// TIA Portal V20 program export: 0 tag tables, 0 data types, 6 data blocks, 13 code blocks (in call order from the OBs), 34 instance data blocks

DATA_BLOCK "DB_Bad_Konfig"   // DB8
{ S7_Optimized_Access := 'TRUE' }
VERSION : 0.5
// stored: AutoNumber true, DBAccessibleFromOPCUA true, DBAccessibleFromWebserver true, IsOnlyStoredInLoadMemory false, IsRetainMemResEnabled false, IsWriteProtectedInAS false, MemoryReserve 100
   VAR
      Bad_Konfig : Array[1.."c_Anzahl_Bad"] of "UDT_Bad_Konfig";
   END_VAR
BEGIN
   Bad_Konfig[7..8].Ausstattung.HatHeizung_1 := TRUE;
   Bad_Konfig[12].Ausstattung.HatHeizung_1 := TRUE;
   Bad_Konfig[25].Ausstattung.HatHeizung_1 := TRUE;
   Bad_Konfig[36].Ausstattung.HatHeizung_1 := TRUE;
   Bad_Konfig[40].Ausstattung.HatHeizung_1 := TRUE;
   Bad_Konfig[46].Ausstattung.HatHeizung_1 := TRUE;
   Bad_Konfig[25].Ausstattung.HatHeizung_2 := TRUE;
   Bad_Konfig[8].Ausstattung.HatPumpe := TRUE;
   Bad_Konfig[12].Ausstattung.HatPumpe := TRUE;
   Bad_Konfig[14].Ausstattung.HatPumpe := TRUE;
   Bad_Konfig[18..19].Ausstattung.HatPumpe := TRUE;
   Bad_Konfig[21].Ausstattung.HatPumpe := TRUE;
   Bad_Konfig[25..26].Ausstattung.HatPumpe := TRUE;
   Bad_Konfig[31].Ausstattung.HatPumpe := TRUE;
   Bad_Konfig[41].Ausstattung.HatPumpe := TRUE;
   Bad_Konfig[45].Ausstattung.HatPumpe := TRUE;
   Bad_Konfig[25].Ausstattung.HatPumpe_FU := TRUE;
   Bad_Konfig[25].Ausstattung.HatWarenbewegung_X := TRUE;
   Bad_Konfig[25].Ausstattung.HatWarenbewegung_Y := TRUE;
   Bad_Konfig[8].Ausstattung.HatUltraschall := TRUE;
   Bad_Konfig[12].Ausstattung.HatUltraschall := TRUE;
   Bad_Konfig[31].Ausstattung.HatGleichrichter := TRUE;
   Bad_Konfig[36].Ausstattung.HatGleichrichter := TRUE;
   Bad_Konfig[40].Ausstattung.HatGleichrichter := TRUE;
   Bad_Konfig[7..8].Ausstattung.HatNiveau := TRUE;
   Bad_Konfig[12].Ausstattung.HatNiveau := TRUE;
   Bad_Konfig[25].Ausstattung.HatNiveau := TRUE;
   Bad_Konfig[36].Ausstattung.HatNiveau := TRUE;
   Bad_Konfig[40].Ausstattung.HatNiveau := TRUE;
   Bad_Konfig[46].Ausstattung.HatNiveau := TRUE;
   Bad_Konfig[1].WT[1..3].Auftragsindex := -1;
   Bad_Konfig[2].WT[1..3].Auftragsindex := -1;
   Bad_Konfig[3].WT[1..3].Auftragsindex := -1;
   Bad_Konfig[4].WT[1..3].Auftragsindex := -1;
   Bad_Konfig[5].WT[1..3].Auftragsindex := -1;
   Bad_Konfig[6].WT[1..3].Auftragsindex := -1;
   Bad_Konfig[7].WT[1..3].Auftragsindex := -1;
   Bad_Konfig[8].WT[1..3].Auftragsindex := -1;
   Bad_Konfig[9].WT[1..3].Auftragsindex := -1;
   Bad_Konfig[10].WT[1..3].Auftragsindex := -1;
   Bad_Konfig[11].WT[1..3].Auftragsindex := -1;
   Bad_Konfig[12].WT[1..3].Auftragsindex := -1;
   Bad_Konfig[13].WT[1..3].Auftragsindex := -1;
   Bad_Konfig[14].WT[1..3].Auftragsindex := -1;
   Bad_Konfig[15].WT[1..3].Auftragsindex := -1;
   Bad_Konfig[16].WT[1..3].Auftragsindex := -1;
   Bad_Konfig[17].WT[1..3].Auftragsindex := -1;
   Bad_Konfig[18].WT[1..3].Auftragsindex := -1;
   Bad_Konfig[19].WT[1..3].Auftragsindex := -1;
   Bad_Konfig[20].WT[1..3].Auftragsindex := -1;
   Bad_Konfig[21].WT[1..3].Auftragsindex := -1;
   Bad_Konfig[22].WT[1..3].Auftragsindex := -1;
   Bad_Konfig[23].WT[1..3].Auftragsindex := -1;
   Bad_Konfig[24].WT[1..3].Auftragsindex := -1;
   Bad_Konfig[25].WT[1..3].Auftragsindex := -1;
   Bad_Konfig[26].WT[1..3].Auftragsindex := -1;
   Bad_Konfig[27].WT[1..3].Auftragsindex := -1;
   Bad_Konfig[28].WT[1..3].Auftragsindex := -1;
   Bad_Konfig[29].WT[1..3].Auftragsindex := -1;
   Bad_Konfig[30].WT[1..3].Auftragsindex := -1;
   Bad_Konfig[31].WT[1..3].Auftragsindex := -1;
   Bad_Konfig[32].WT[1..3].Auftragsindex := -1;
   Bad_Konfig[33].WT[1..3].Auftragsindex := -1;
   Bad_Konfig[34].WT[1..3].Auftragsindex := -1;
   Bad_Konfig[35].WT[1..3].Auftragsindex := -1;
   Bad_Konfig[36].WT[1..3].Auftragsindex := -1;
   Bad_Konfig[37].WT[1..3].Auftragsindex := -1;
   Bad_Konfig[38].WT[1..3].Auftragsindex := -1;
   Bad_Konfig[39].WT[1..3].Auftragsindex := -1;
   Bad_Konfig[40].WT[1..3].Auftragsindex := -1;
   Bad_Konfig[41].WT[1..3].Auftragsindex := -1;
   Bad_Konfig[42].WT[1..3].Auftragsindex := -1;
   Bad_Konfig[43].WT[1..3].Auftragsindex := -1;
   Bad_Konfig[44].WT[1..3].Auftragsindex := -1;
   Bad_Konfig[45].WT[1..3].Auftragsindex := -1;
   Bad_Konfig[46].WT[1..3].Auftragsindex := -1;
   Bad_Konfig[47].WT[1..3].Auftragsindex := -1;
   Bad_Konfig[1].WT[1..3].SchrittIndex := -1;
   Bad_Konfig[2].WT[1..3].SchrittIndex := -1;
   Bad_Konfig[3].WT[1..3].SchrittIndex := -1;
   Bad_Konfig[4].WT[1..3].SchrittIndex := -1;
   Bad_Konfig[5].WT[1..3].SchrittIndex := -1;
   Bad_Konfig[6].WT[1..3].SchrittIndex := -1;
   Bad_Konfig[7].WT[1..3].SchrittIndex := -1;
   Bad_Konfig[8].WT[1..3].SchrittIndex := -1;
   Bad_Konfig[9].WT[1..3].SchrittIndex := -1;
   Bad_Konfig[10].WT[1..3].SchrittIndex := -1;
   Bad_Konfig[11].WT[1..3].SchrittIndex := -1;
   Bad_Konfig[12].WT[1..3].SchrittIndex := -1;
   Bad_Konfig[13].WT[1..3].SchrittIndex := -1;
   Bad_Konfig[14].WT[1..3].SchrittIndex := -1;
   Bad_Konfig[15].WT[1..3].SchrittIndex := -1;
   Bad_Konfig[16].WT[1..3].SchrittIndex := -1;
   Bad_Konfig[17].WT[1..3].SchrittIndex := -1;
   Bad_Konfig[18].WT[1..3].SchrittIndex := -1;
   Bad_Konfig[19].WT[1..3].SchrittIndex := -1;
   Bad_Konfig[20].WT[1..3].SchrittIndex := -1;
   Bad_Konfig[21].WT[1..3].SchrittIndex := -1;
   Bad_Konfig[22].WT[1..3].SchrittIndex := -1;
   Bad_Konfig[23].WT[1..3].SchrittIndex := -1;
   Bad_Konfig[24].WT[1..3].SchrittIndex := -1;
   Bad_Konfig[25].WT[1..3].SchrittIndex := -1;
   Bad_Konfig[26].WT[1..3].SchrittIndex := -1;
   Bad_Konfig[27].WT[1..3].SchrittIndex := -1;
   Bad_Konfig[28].WT[1..3].SchrittIndex := -1;
   Bad_Konfig[29].WT[1..3].SchrittIndex := -1;
   Bad_Konfig[30].WT[1..3].SchrittIndex := -1;
   Bad_Konfig[31].WT[1..3].SchrittIndex := -1;
   Bad_Konfig[32].WT[1..3].SchrittIndex := -1;
   Bad_Konfig[33].WT[1..3].SchrittIndex := -1;
   Bad_Konfig[34].WT[1..3].SchrittIndex := -1;
   Bad_Konfig[35].WT[1..3].SchrittIndex := -1;
   Bad_Konfig[36].WT[1..3].SchrittIndex := -1;
   Bad_Konfig[37].WT[1..3].SchrittIndex := -1;
   Bad_Konfig[38].WT[1..3].SchrittIndex := -1;
   Bad_Konfig[39].WT[1..3].SchrittIndex := -1;
   Bad_Konfig[40].WT[1..3].SchrittIndex := -1;
   Bad_Konfig[41].WT[1..3].SchrittIndex := -1;
   Bad_Konfig[42].WT[1..3].SchrittIndex := -1;
   Bad_Konfig[43].WT[1..3].SchrittIndex := -1;
   Bad_Konfig[44].WT[1..3].SchrittIndex := -1;
   Bad_Konfig[45].WT[1..3].SchrittIndex := -1;
   Bad_Konfig[46].WT[1..3].SchrittIndex := -1;
   Bad_Konfig[47].WT[1..3].SchrittIndex := -1;
END_DATA_BLOCK

DATA_BLOCK "DB_HMI"   // DB4
{ S7_Optimized_Access := 'TRUE' }
VERSION : 0.1
// stored: AutoNumber true, DBAccessibleFromOPCUA true, DBAccessibleFromWebserver true, IsOnlyStoredInLoadMemory false, IsRetainMemResEnabled false, IsWriteProtectedInAS false, MemoryReserve 100
   VAR
      Benutzerverwaltung_User_Daten { S7_SetPoint := 'True'} : "UDT_Benutzer";
      Benutzerverwaltung_User_create { S7_SetPoint := 'True'} : Bool;
      Benutzerverwaltung_User_update : Bool;
      Benutzerverwaltung_User_delete : Bool;
      Benutzerverwaltung_Freigaben_Prozessgruppen_User_change : Bool;
      Benutzerverwaltung_Status : Int;
      Benutzerverwaltung_Freigabe_Prozessgruppen_User_ID_ausgewählt : Int;
      Benutzerverwaltung_Freigabe_Prozessgruppen_Prozessgruppen : Array[1.."c_Prozessgruppen"] of Bool;
      Benutzerverwaltung_Login_Name : String;
      Benutzerverwaltung_Login_Passwort : String;
      Benutzerverwaltung_Login_Loginbutton : Bool;
      Benutzerverwaltung_Login_Logoutbutton : Bool;
      Benutzerverwaltung_Login_Login_Ok : Bool;
      Prozessparameter_Status : Int;
      Prozessparameter_Prozessgruppen_save : Bool;
      Prozessparameter_Prozessgruppen_Prozessgruppe : "UDT_Prozessgruppen";
      Prozessparameter_Artikel_add { S7_SetPoint := 'True'} : "UDT_Artikel";
      Prozessparameter_Artikel_save { S7_SetPoint := 'True'} : Bool;
      Prozessparameter_Artikel_delete : Bool;
      Prozessparameter_Artikel_assign : Bool;
      Prozessparameter_Artikel_remove : Bool;
      "Prozessparameter_Prozessgruppe_ID_assign/remove" : Int;
      "Prozessparameter_Artikel_ID_assign/remove" : Int;
      Angewähltes_Bad : USInt;
      Handbetrieb { S7_SetPoint := 'True'} : "UDT_Handbetrieb";
   END_VAR
BEGIN
END_DATA_BLOCK

DATA_BLOCK "DB_CPU_to_IPC"   // DB3
{ S7_Optimized_Access := 'TRUE' }
VERSION : 0.2
// stored: AutoNumber true, DBAccessibleFromOPCUA true, DBAccessibleFromWebserver true, IsOnlyStoredInLoadMemory false, IsRetainMemResEnabled false, IsWriteProtectedInAS false, MemoryReserve 100
   VAR
      Bad : Array[1.."c_Anzahl_Bad"] of "UDT_Bad_Rueckmeldung";
      Not_Halt_Aktiv : Bool;
      Not_Aus_OK : Bool;
      Auftrag_Abgeschlossen : Array[0..9] of Bool;
   END_VAR
BEGIN
END_DATA_BLOCK

DATA_BLOCK "DB_Fehlermeldungen"   // DB39
{ S7_Optimized_Access := 'TRUE' }
VERSION : 0.2
// FI-Schutz ausgeloest (Heizungen)
// stored: AutoNumber true, DBAccessibleFromOPCUA true, DBAccessibleFromWebserver true, IsOnlyStoredInLoadMemory false, IsRetainMemResEnabled false, IsWriteProtectedInAS false, MemoryReserve 100
   VAR
      FI_Heizung_Bad_7 : Bool;   // 1 - FI-Schutz 200F1 Heizung Bad 7 ausgeloest
      FI_Heizung_Bad_8 : Bool;   // 2 - FI-Schutz 210F1 Heizung Bad 8 ausgeloest
      FI_Heizung_Bad_12 : Bool;   // 3 - FI-Schutz 220F1 Heizung Bad 12 ausgeloest
      FI_Heizung_Bad_25 : Bool;   // 4 - FI+Motorschutz 270/271 Heizung Bad 25 ausgeloest
      FI_Heizung_Bad_36 : Bool;   // 5 - FI-Schutz 300F1 Heizung Bad 36 ausgeloest
      FI_Heizung_Bad_40 : Bool;   // 6 - FI-Schutz 310F1 Heizung Bad 40 ausgeloest
      FI_Heizung_Bad_46 : Bool;   // 7 - FI-Schutz 340F1 Heizung Bad 46 ausgeloest Uebertemperatur (Heizungen)
      Uebertemp_Bad_7 : Bool;   // 8 - Uebertemperatur Heizung Bad 7
      Uebertemp_Bad_8 : Bool;   // 9 - Uebertemperatur Heizung Bad 8
      Uebertemp_Bad_12 : Bool;   // 10 - Uebertemperatur Heizung Bad 12
      Uebertemp_Bad_25 : Bool;   // 11 - Uebertemperatur Heizung Bad 25
      Uebertemp_Bad_36 : Bool;   // 12 - Uebertemperatur Heizung Bad 36
      Uebertemp_Bad_40 : Bool;   // 13 - Uebertemperatur Heizung Bad 40
      Uebertemp_Bad_46 : Bool;   // 14 - Uebertemperatur Heizung Bad 46 Motorschutz Pumpe ausgeloest
      Motorschutz_Pumpe_Bad_8 : Bool;   // 15 - Motorschutz 215Q1 Pumpe Bad 8 ausgeloest
      Motorschutz_Pumpe_Bad_12 : Bool;   // 16 - Motorschutz 225Q1 Pumpe Bad 12 ausgeloest
      Motorschutz_Pumpe_Bad_14 : Bool;   // 17 - Motorschutz 235Q1 Pumpe Bad 14 ausgeloest
      Motorschutz_Pumpe_Bad_18 : Bool;   // 18 - Motorschutz 245Q1 Pumpe Bad 18 ausgeloest
      Motorschutz_Pumpe_Bad_19 : Bool;   // 19 - Motorschutz 255Q1 Pumpe Bad 19 ausgeloest
      Motorschutz_Pumpe_Bad_21 : Bool;   // 20 - Motorschutz 265Q1 Pumpe Bad 21 ausgeloest
      Motorschutz_Pumpe_Bad_25 : Bool;   // 21 - Motorschutz 275Q1 Pumpe Bad 25 ausgeloest
      Motorschutz_Pumpe_Bad_26 : Bool;   // 22 - Motorschutz 285Q1 Pumpe Bad 26 ausgeloest
      Motorschutz_Pumpe_Bad_31 : Bool;   // 23 - Motorschutz 295Q1 Pumpe Bad 31 ausgeloest
      Motorschutz_Pumpe_Bad_41 : Bool;   // 24 - Motorschutz 325Q1 Pumpe Bad 41 ausgeloest
      Motorschutz_Pumpe_Bad_45 : Bool;   // 25 - Motorschutz 335Q1 Pumpe Bad 45 ausgeloest Wartungsschalter Pumpe nicht eingeschaltet
      Wartungsschalter_Pumpe_Bad_8 : Bool;   // 26 - Wartungsschalter Pumpe Bad 8 nicht eingeschaltet
      Wartungsschalter_Pumpe_Bad_12 : Bool;   // 27 - Wartungsschalter Pumpe Bad 12 nicht eingeschaltet
      Wartungsschalter_Pumpe_Bad_14 : Bool;   // 28 - Wartungsschalter Pumpe Bad 14 nicht eingeschaltet
      Wartungsschalter_Pumpe_Bad_18 : Bool;   // 29 - Wartungsschalter Pumpe Bad 18 nicht eingeschaltet
      Wartungsschalter_Pumpe_Bad_19 : Bool;   // 30 - Wartungsschalter Pumpe Bad 19 nicht eingeschaltet
      Wartungsschalter_Pumpe_Bad_21 : Bool;   // 31 - Wartungsschalter Pumpe Bad 21 nicht eingeschaltet
      Wartungsschalter_Pumpe_Bad_25 : Bool;   // 32 - Wartungsschalter Pumpe Bad 25 nicht eingeschaltet
      Wartungsschalter_Pumpe_Bad_26 : Bool;   // 33 - Wartungsschalter Pumpe Bad 26 nicht eingeschaltet
      Wartungsschalter_Pumpe_Bad_31 : Bool;   // 34 - Wartungsschalter Pumpe Bad 31 nicht eingeschaltet
      Wartungsschalter_Pumpe_Bad_41 : Bool;   // 35 - Wartungsschalter Pumpe Bad 41 nicht eingeschaltet
      Wartungsschalter_Pumpe_Bad_45 : Bool;   // 36 - Wartungsschalter Pumpe Bad 45 nicht eingeschaltet Niveau nicht OK
      Niveau_Bad_7 : Bool;   // 37 - Niveau Bad 7 nicht OK
      Niveau_Bad_8 : Bool;   // 38 - Niveau Bad 8 nicht OK
      Niveau_Bad_12 : Bool;   // 39 - Niveau Bad 12 nicht OK
      Niveau_Bad_25 : Bool;   // 40 - Niveau Bad 25 nicht OK
      Niveau_Bad_36 : Bool;   // 41 - Niveau Bad 36 nicht OK
      Niveau_Bad_40 : Bool;   // 42 - Niveau Bad 40 nicht OK
      Niveau_Bad_46 : Bool;   // 43 - Niveau Bad 46 nicht OK Frequenzumrichter Stoerung (angesteuert aber nicht bereit, 3s verzoegert)
      FU_Pumpe_Bad_25 : Bool;   // 44 - FU Umwaelzpumpe Bad 25 Stoerung
      FU_WB1_Bad_25 : Bool;   // 45 - FU Warenbewegung 1 Bad 25 Stoerung
      FU_WB2_Bad_25 : Bool;   // 46 - FU Warenbewegung 2 Bad 25 Stoerung Motorschutz Warenbewegung ausgeloest
      Motorschutz_WB1_Bad_25 : Bool;   // 47 - Motorschutz 276Q1 Warenbewegung 1 Bad 25 ausgeloest
      Motorschutz_WB2_Bad_25 : Bool;   // 48 - Motorschutz 277Q1 Warenbewegung 2 Bad 25 ausgeloest PT100 Sensorstoerung (Drahtbruch oder Kurzschluss)
      PT100_Bad_7 : Bool;   // 49 - PT100 Heizung Bad 7 Sensorstoerung
      PT100_Bad_8 : Bool;   // 50 - PT100 Heizung Bad 8 Sensorstoerung
      PT100_Bad_12 : Bool;   // 51 - PT100 Heizung Bad 12 Sensorstoerung
      PT100_Bad_25_H1 : Bool;   // 52 - PT100 Heizung 1 Bad 25 Sensorstoerung
      PT100_Bad_25_H2 : Bool;   // 53 - PT100 Heizung 2 Bad 25 Sensorstoerung
      PT100_Bad_36 : Bool;   // 54 - PT100 Heizung Bad 36 Sensorstoerung
      PT100_Bad_40 : Bool;   // 55 - PT100 Heizung Bad 40 Sensorstoerung
      PT100_Bad_46 : Bool;   // 56 - PT100 Heizung Bad 46 Sensorstoerung Walchem Controller
      Fehler_Walchem_Controller : Bool;   // 57 - Alarm Walchem Controller Bad 25 Not-Halt
      Not_Halt : Bool;   // 58 - Not-Halt ausgeloest
   END_VAR
BEGIN
END_DATA_BLOCK

DATA_BLOCK "DB_FlexKraft_Data"   // DB5
{ S7_Optimized_Access := 'FALSE' }
VERSION : 0.1
// ==============================================================================
//  DB: Daten aller drei FlexKraft-GerÃ¤te
// ==============================================================================
// stored: AutoNumber true, DBAccessibleFromOPCUA true, DBAccessibleFromWebserver true, IsOnlyStoredInLoadMemory false, IsWriteProtectedInAS false
   VAR
      FK_1 { S7_SetPoint := 'True'} : "UDT_FlexKraft_Device";   // ModbusAdr 2 (Gateway-Bytes 0..31)
      FK_2 { S7_SetPoint := 'True'} : "UDT_FlexKraft_Device";   // ModbusAdr 3 (Gateway-Bytes 32..63)
      FK_3 { S7_SetPoint := 'True'} : "UDT_FlexKraft_Device";   // ModbusAdr 4 (Gateway-Bytes 64..95)
   END_VAR
BEGIN
END_DATA_BLOCK

DATA_BLOCK "DB_IPC_to_CPU"   // DB2
{ S7_Optimized_Access := 'TRUE' }
VERSION : 0.1
// stored: AutoNumber true, DBAccessibleFromOPCUA true, DBAccessibleFromWebserver true, IsOnlyStoredInLoadMemory false, IsRetainMemResEnabled false, IsWriteProtectedInAS false, MemoryReserve 100
   VAR
      Auftrag : Array[0..9] of "UDT_Prozessroute";
      Handbetrieb : Array[1.."c_Anzahl_Bad"] of "UDT_Handbetrieb";
      Not_Halt_Reset : Bool;
      Lampentest : Bool;   // Virtuelle Tasten fuer Baeder ohne KP8 (Bad 2, 20, 47)
      Virtuelle_Tasten : Struct
         Bad_2 : Struct
            WT_Einsetzen : Array[1..3] of Bool;
            WT_Entnehmen : Array[1..3] of Bool;
         END_STRUCT;
         Bad_20 : Struct
            WT_Einsetzen : Array[1..3] of Bool;
            WT_Entnehmen : Array[1..3] of Bool;
         END_STRUCT;
         Bad_47 : Struct
            WT_Einsetzen : Array[1..3] of Bool;
            WT_Entnehmen : Array[1..3] of Bool;   // Leerlauf-Parameter pro Bad (Zustand 1: betriebsbereit halten)
         END_STRUCT;
      END_STRUCT;
   END_VAR
   VAR RETAIN
      Leerlauf : Array[1.."c_Anzahl_Bad"] of "UDT_Peripherie_Soll";   // Standby-Parameter pro Bad (Zustand 2: abgesenkt, Energie sparen)
      Standby : Array[1.."c_Anzahl_Bad"] of "UDT_Peripherie_Soll";   // Anlagenzustand: 0=undefiniert/alles aus, 1=Leerlauf, 2=Standby
   END_VAR
   VAR
      Zustand : Array[1.."c_Anzahl_Bad"] of Int;   // PT100 Offset pro Bad (vom IPC einstellbar, in Grad Celsius)
      PT100_Offset : Array[1.."c_Anzahl_Bad"] of Real;
   END_VAR
BEGIN
   PT100_Offset[7] := -4.0;
   PT100_Offset[8] := -3.8;
   PT100_Offset[12] := -4.0;
   PT100_Offset[25] := -5.8;
   PT100_Offset[36] := -3.4;
   PT100_Offset[40] := -3.2;
   PT100_Offset[46] := -3.0;
END_DATA_BLOCK

ORGANIZATION_BLOCK "Main"   // OB1, LAD, ProgramCycle
TITLE = "Main Program Sweep (Cycle)"
{ S7_Optimized_Access := 'TRUE' }
VERSION : 0.1
// stored: AutoNumber true, IsIECCheckEnabled false, SetENOAutomatically false
   VAR_INPUT
      Initial_Call : Bool;   // Initial call of this OB
      Remanence : Bool;   // =True, if remanent data are available
   END_VAR
   VAR_TEMP
      Lampentest_Ein : Bool;
      Blinktakt : Bool;
   END_VAR
BEGIN

REGION Network 1 (SCL): Eingaenge Lesen
   //KP8_1
   "FB_KP8_DB_1".KP8.Rohdaten.IB_Tasten := "KP8_1_IB_Tasten";
   "FB_KP8_DB_1".KP8.Rohdaten.IB_DI := "KP8_1_IB_DI";
   "FB_KP8_DB_1"();

   //KP8_2
   "FB_KP8_DB_2".KP8.Rohdaten.IB_Tasten := "KP8_2_IB_Tasten";
   "FB_KP8_DB_2".KP8.Rohdaten.IB_DI := "KP8_2_IB_DI";
   "FB_KP8_DB_2"();

   //KP8_3
   "FB_KP8_DB_3".KP8.Rohdaten.IB_Tasten := "KP8_3_IB_Tasten";
   "FB_KP8_DB_3".KP8.Rohdaten.IB_DI := "KP8_3_IB_DI";
   "FB_KP8_DB_3"();

   //KP8_4
   "FB_KP8_DB_4".KP8.Rohdaten.IB_Tasten := "KP8_4_IB_Tasten";
   "FB_KP8_DB_4".KP8.Rohdaten.IB_DI := "KP8_4_IB_DI";
   "FB_KP8_DB_4"();

   //KP8_5
   "FB_KP8_DB_5".KP8.Rohdaten.IB_Tasten := "KP8_5_IB_Tasten";
   "FB_KP8_DB_5".KP8.Rohdaten.IB_DI := "KP8_5_IB_DI";
   "FB_KP8_DB_5"();

   //KP8_6
   "FB_KP8_DB_6".KP8.Rohdaten.IB_Tasten := "KP8_6_IB_Tasten";
   "FB_KP8_DB_6".KP8.Rohdaten.IB_DI := "KP8_6_IB_DI";
   "FB_KP8_DB_6"();

   //KP8_7
   "FB_KP8_DB_7".KP8.Rohdaten.IB_Tasten := "KP8_7_IB_Tasten";
   "FB_KP8_DB_7".KP8.Rohdaten.IB_DI := "KP8_7_IB_DI";
   "FB_KP8_DB_7"();

   //KP8_8
   "FB_KP8_DB_8".KP8.Rohdaten.IB_Tasten := "KP8_8_IB_Tasten";
   "FB_KP8_DB_8".KP8.Rohdaten.IB_DI := "KP8_8_IB_DI";
   "FB_KP8_DB_8"();

   //KP8_9
   "FB_KP8_DB_9".KP8.Rohdaten.IB_Tasten := "KP8_9_IB_Tasten";
   "FB_KP8_DB_9".KP8.Rohdaten.IB_DI := "KP8_9_IB_DI";
   "FB_KP8_DB_9"();

   //KP8_10
   "FB_KP8_DB_10".KP8.Rohdaten.IB_Tasten := "KP8_10_IB_Tasten";
   "FB_KP8_DB_10".KP8.Rohdaten.IB_DI := "KP8_10_IB_DI";
   "FB_KP8_DB_10"();

   //KP8_11
   "FB_KP8_DB_11".KP8.Rohdaten.IB_Tasten := "KP8_11_IB_Tasten";
   "FB_KP8_DB_11".KP8.Rohdaten.IB_DI := "KP8_11_IB_DI";
   "FB_KP8_DB_11"();

   //KP8_12
   "FB_KP8_DB_12".KP8.Rohdaten.IB_Tasten := "KP8_12_IB_Tasten";
   "FB_KP8_DB_12".KP8.Rohdaten.IB_DI := "KP8_12_IB_DI";
   "FB_KP8_DB_12"();

   //KP8_13
   "FB_KP8_DB_13".KP8.Rohdaten.IB_Tasten := "KP8_13_IB_Tasten";
   "FB_KP8_DB_13".KP8.Rohdaten.IB_DI := "KP8_13_IB_DI";
   "FB_KP8_DB_13"();

   //KP8_14
   "FB_KP8_DB_14".KP8.Rohdaten.IB_Tasten := "KP8_14_IB_Tasten";
   "FB_KP8_DB_14".KP8.Rohdaten.IB_DI := "KP8_14_IB_DI";
   "FB_KP8_DB_14"();

   //KP8_15
   "FB_KP8_DB_15".KP8.Rohdaten.IB_Tasten := "KP8_15_IB_Tasten";
   "FB_KP8_DB_15".KP8.Rohdaten.IB_DI := "KP8_15_IB_DI";
   "FB_KP8_DB_15"();

   //KP8_16
   "FB_KP8_DB_16".KP8.Rohdaten.IB_Tasten := "KP8_16_IB_Tasten";
   "FB_KP8_DB_16".KP8.Rohdaten.IB_DI := "KP8_16_IB_DI";
   "FB_KP8_DB_16"();

   //KP8_17
   "FB_KP8_DB_17".KP8.Rohdaten.IB_Tasten := "KP8_17_IB_Tasten";
   "FB_KP8_DB_17".KP8.Rohdaten.IB_DI := "KP8_17_IB_DI";
   "FB_KP8_DB_17"();

   //KP8_18
   "FB_KP8_DB_18".KP8.Rohdaten.IB_Tasten := "KP8_18_IB_Tasten";
   "FB_KP8_DB_18".KP8.Rohdaten.IB_DI := "KP8_18_IB_DI";
   "FB_KP8_DB_18"();

   //KP8_19
   "FB_KP8_DB_19".KP8.Rohdaten.IB_Tasten := "KP8_19_IB_Tasten";
   "FB_KP8_DB_19".KP8.Rohdaten.IB_DI := "KP8_19_IB_DI";
   "FB_KP8_DB_19"();

   //KP8_20
   "FB_KP8_DB_20".KP8.Rohdaten.IB_Tasten := "KP8_20_IB_Tasten";
   "FB_KP8_DB_20".KP8.Rohdaten.IB_DI := "KP8_20_IB_DI";
   "FB_KP8_DB_20"();

   //KP8_21
   "FB_KP8_DB_21".KP8.Rohdaten.IB_Tasten := "KP8_21_IB_Tasten";
   "FB_KP8_DB_21".KP8.Rohdaten.IB_DI := "KP8_21_IB_DI";
   "FB_KP8_DB_21"();

   //KP8_22
   "FB_KP8_DB_22".KP8.Rohdaten.IB_Tasten := "KP8_22_IB_Tasten";
   "FB_KP8_DB_22".KP8.Rohdaten.IB_DI := "KP8_22_IB_DI";
   "FB_KP8_DB_22"();

   //KP8_23
   "FB_KP8_DB_23".KP8.Rohdaten.IB_Tasten := "KP8_23_IB_Tasten";
   "FB_KP8_DB_23".KP8.Rohdaten.IB_DI := "KP8_23_IB_DI";
   "FB_KP8_DB_23"();

   //KP8_24
   "FB_KP8_DB_24".KP8.Rohdaten.IB_Tasten := "KP8_24_IB_Tasten";
   "FB_KP8_DB_24".KP8.Rohdaten.IB_DI := "KP8_24_IB_DI";
   "FB_KP8_DB_24"();

   //KP8_25
   "FB_KP8_DB_25".KP8.Rohdaten.IB_Tasten := "KP8_25_IB_Tasten";
   "FB_KP8_DB_25".KP8.Rohdaten.IB_DI := "KP8_25_IB_DI";
   "FB_KP8_DB_25"();

   //KP8_26
   "FB_KP8_DB_26".KP8.Rohdaten.IB_Tasten := "KP8_26_IB_Tasten";
   "FB_KP8_DB_26".KP8.Rohdaten.IB_DI := "KP8_26_IB_DI";
   "FB_KP8_DB_26"();

   //KP8_27
   "FB_KP8_DB_27".KP8.Rohdaten.IB_Tasten := "KP8_27_IB_Tasten";
   "FB_KP8_DB_27".KP8.Rohdaten.IB_DI := "KP8_27_IB_DI";
   "FB_KP8_DB_27"();

   //KP8_28
   "FB_KP8_DB_28".KP8.Rohdaten.IB_Tasten := "KP8_28_IB_Tasten";
   "FB_KP8_DB_28".KP8.Rohdaten.IB_DI := "KP8_28_IB_DI";
   "FB_KP8_DB_28"();
END_REGION

REGION Network 2 (SCL): Badlogik
   "FB_Anlagensteuerung_DB"(Blink_Takt:="Clock_1Hz",
                            Clock_10Hz:="Clock_10Hz",
                            Not_Halt_Aktiv:=NOT "Not-Aus ist OK");
END_REGION

REGION Network 3 (SCL): Flexkraft
   // ----- 1) Eingänge aus Peripherie in den DB kopieren -----

   // FK_1 (IB500..IB531)
   "DB_FlexKraft_Data".FK_1.In.Reserved0            := "Flexkraft_1";    //IW500
   "DB_FlexKraft_Data".FK_1.In.StatusRegister       := "Flexkraft_2";    //IW502
   "DB_FlexKraft_Data".FK_1.In.WarningsRegister     := "Flexkraft_3";    //IW504
   "DB_FlexKraft_Data".FK_1.In.AlarmsRegister       := "Flexkraft_4";    //IW506
   "DB_FlexKraft_Data".FK_1.In.OutputVoltage        := "Flexkraft_5";    //IW508
   "DB_FlexKraft_Data".FK_1.In.OutputCurrent        := "Flexkraft_6";    //IW510
   "DB_FlexKraft_Data".FK_1.In.ProcessTime_HW       := "Flexkraft_7";    //IW512
   "DB_FlexKraft_Data".FK_1.In.ProcessTime_LW       := "Flexkraft_8";    //IW514
   "DB_FlexKraft_Data".FK_1.In.Ah_HW                := "Flexkraft_9";    //IW516
   "DB_FlexKraft_Data".FK_1.In.Ah_LW                := "Flexkraft_10";   //IW518

   // FK_2 (IB532..IB563)
   "DB_FlexKraft_Data".FK_2.In.Reserved0           := "Flexkraft_20";    //IW532
   "DB_FlexKraft_Data".FK_2.In.StatusRegister      := "Flexkraft_21";    //IW534
   "DB_FlexKraft_Data".FK_2.In.WarningsRegister    := "Flexkraft_22";    //IW536
   "DB_FlexKraft_Data".FK_2.In.AlarmsRegister      := "Flexkraft_23";    //IW538
   "DB_FlexKraft_Data".FK_2.In.OutputVoltage       := "Flexkraft_24";    //IW540
   "DB_FlexKraft_Data".FK_2.In.OutputCurrent       := "Flexkraft_25";    //IW542
   "DB_FlexKraft_Data".FK_2.In.ProcessTime_HW      := "Flexkraft_26";    //IW544
   "DB_FlexKraft_Data".FK_2.In.ProcessTime_LW      := "Flexkraft_27";    //IW546
   "DB_FlexKraft_Data".FK_2.In.Ah_HW               := "Flexkraft_28";    //IW548
   "DB_FlexKraft_Data".FK_2.In.Ah_LW               := "Flexkraft_29";    //IW550

   // FK_3 (IB564..IB595)
   "DB_FlexKraft_Data".FK_3.In.Reserved0           := "Flexkraft_30";    //IW564
   "DB_FlexKraft_Data".FK_3.In.StatusRegister      := "Flexkraft_31";    //IW566
   "DB_FlexKraft_Data".FK_3.In.WarningsRegister    := "Flexkraft_32";    //IW568
   "DB_FlexKraft_Data".FK_3.In.AlarmsRegister      := "Flexkraft_33";    //IW570
   "DB_FlexKraft_Data".FK_3.In.OutputVoltage       := "Flexkraft_34";    //IW572
   "DB_FlexKraft_Data".FK_3.In.OutputCurrent       := "Flexkraft_35";    //IW574
   "DB_FlexKraft_Data".FK_3.In.ProcessTime_HW      := "Flexkraft_36";    //IW576
   "DB_FlexKraft_Data".FK_3.In.ProcessTime_LW      := "Flexkraft_37";    //IW578
   "DB_FlexKraft_Data".FK_3.In.Ah_HW               := "Flexkraft_38";    //IW580
   "DB_FlexKraft_Data".FK_3.In.Ah_LW               := "Flexkraft_39";    //IW582

   // ----- 2) FB-Aufruf (1 Instanz pro Gerät) -----
   "FB_FlexKraft_DB"(bOn:="DB_Bad_Konfig".Bad_Konfig[40].GR_Aktiv,
                     bStartA:="DB_Bad_Konfig".Bad_Konfig[40].GR_Aktiv,
                     iSetVoltage_cV:="DB_Bad_Konfig".Bad_Konfig[40].GR_Spannung_Soll * 100,
                     iSetCurrent_raw:="DB_Bad_Konfig".Bad_Konfig[40].GR_Strom_Soll,
                     stDev:="DB_FlexKraft_Data".FK_1);

   "FB_FlexKraft_DB_1"(bOn:="DB_Bad_Konfig".Bad_Konfig[36].GR_Aktiv,
                       bStartA:="DB_Bad_Konfig".Bad_Konfig[36].GR_Aktiv,
                       iSetVoltage_cV:="DB_Bad_Konfig".Bad_Konfig[36].GR_Spannung_Soll * 100,
                       iSetCurrent_raw:="DB_Bad_Konfig".Bad_Konfig[36].GR_Strom_Soll,
                       stDev:="DB_FlexKraft_Data".FK_2);

   "FB_FlexKraft_DB_2"(bOn:="DB_Bad_Konfig".Bad_Konfig[31].GR_Aktiv,
                       bStartA:="DB_Bad_Konfig".Bad_Konfig[31].GR_Aktiv,
                       iSetVoltage_cV:="DB_Bad_Konfig".Bad_Konfig[31].GR_Spannung_Soll * 100,
                       iSetCurrent_raw:="DB_Bad_Konfig".Bad_Konfig[31].GR_Strom_Soll,
                       stDev:="DB_FlexKraft_Data".FK_3);


   // ----- 3) Ausgänge aus dem DB in die Peripherie kopieren -----

   // FK_1 (QB500..QB531)
   "Flexkraft_11"    := "DB_FlexKraft_Data".FK_1.Out.PageNo;                 //QW500
   "Flexkraft_12"    := "DB_FlexKraft_Data".FK_1.Out.ControlRegister;        //QW502
   "Flexkraft_13"    := "DB_FlexKraft_Data".FK_1.Out.SetVoltage;             //QW504
   "Flexkraft_14"    := "DB_FlexKraft_Data".FK_1.Out.SetCurrent;             //QW506
   "Flexkraft_15"    := "DB_FlexKraft_Data".FK_1.Out.ProcessTimerLimit_HW;   //QW508
   "Flexkraft_16"    := "DB_FlexKraft_Data".FK_1.Out.ProcessTimerLimit_LW;   //QW510
   "Flexkraft_17"    := "DB_FlexKraft_Data".FK_1.Out.AhLimit_HW;             //QW512
   "Flexkraft_18"    := "DB_FlexKraft_Data".FK_1.Out.AhLimit_LW;             //QW514
   "Flexkraft_19"    := "DB_FlexKraft_Data".FK_1.Out.Startramp;              //QW516

   // FK_2 (QB532..QB563)
   "Flexkraft_40"    :="DB_FlexKraft_Data".FK_2.Out.PageNo;                  //QW532
   "Flexkraft_41"    :="DB_FlexKraft_Data".FK_2.Out.ControlRegister;         //QW534
   "Flexkraft_42"    :="DB_FlexKraft_Data".FK_2.Out.SetVoltage;              //QW536
   "Flexkraft_43"    :="DB_FlexKraft_Data".FK_2.Out.SetCurrent;              //QW538
   "Flexkraft_44"    :="DB_FlexKraft_Data".FK_2.Out.ProcessTimerLimit_HW;    //QW540
   "Flexkraft_45"    :="DB_FlexKraft_Data".FK_2.Out.ProcessTimerLimit_LW;    //QW542
   "Flexkraft_46"    :="DB_FlexKraft_Data".FK_2.Out.AhLimit_HW;              //QW544
   "Flexkraft_49"    :="DB_FlexKraft_Data".FK_2.Out.AhLimit_LW;              //QW546
   "Flexkraft_48"    :="DB_FlexKraft_Data".FK_2.Out.Startramp;               //QW548

   // FK_3 (QB564..QB595)
   "Flexkraft_47"    :="DB_FlexKraft_Data".FK_3.Out.PageNo;                  //QW564
   "Flexkraft_50"    :="DB_FlexKraft_Data".FK_3.Out.ControlRegister;         //QW566
   "Flexkraft_51"    :="DB_FlexKraft_Data".FK_3.Out.SetVoltage;              //QW568
   "Flexkraft_52"    :="DB_FlexKraft_Data".FK_3.Out.SetCurrent;              //QW570
   "Flexkraft_54"    :="DB_FlexKraft_Data".FK_3.Out.ProcessTimerLimit_HW;    //QW572
   "Flexkraft_53"    :="DB_FlexKraft_Data".FK_3.Out.ProcessTimerLimit_LW;    //QW574
   "Flexkraft_55"    :="DB_FlexKraft_Data".FK_3.Out.AhLimit_HW;              //QW576
   "Flexkraft_56"    :="DB_FlexKraft_Data".FK_3.Out.AhLimit_LW;              //QW578
   "Flexkraft_57"    :="DB_FlexKraft_Data".FK_3.Out.Startramp;               //QW580
END_REGION

REGION Network 4 (SCL): Ausgaenge schreiben

   //KP8_1
   "FB_KP8_DB_1"();
   "KP8_1_QB_Rot" := "FB_KP8_DB_1".KP8.Rohdaten.QB_Rot;
   "KP8_1_QB_Gruen" := "FB_KP8_DB_1".KP8.Rohdaten.QB_Gruen;
   "KP8_1_QB_Blau" := "FB_KP8_DB_1".KP8.Rohdaten.QB_Blau;
   "KP8_1_QB_DO" := "FB_KP8_DB_1".KP8.Rohdaten.QB_DO;

   //KP8_2
   "FB_KP8_DB_2"();
   "KP8_2_QB_Rot" := "FB_KP8_DB_2".KP8.Rohdaten.QB_Rot;
   "KP8_2_QB_Gruen" := "FB_KP8_DB_2".KP8.Rohdaten.QB_Gruen;
   "KP8_2_QB_Blau" := "FB_KP8_DB_2".KP8.Rohdaten.QB_Blau;
   "KP8_2_QB_DO" := "FB_KP8_DB_2".KP8.Rohdaten.QB_DO;

   //KP8_3
   "FB_KP8_DB_3"();
   "KP8_3_QB_Rot" := "FB_KP8_DB_3".KP8.Rohdaten.QB_Rot;
   "KP8_3_QB_Gruen" := "FB_KP8_DB_3".KP8.Rohdaten.QB_Gruen;
   "KP8_3_QB_Blau" := "FB_KP8_DB_3".KP8.Rohdaten.QB_Blau;
   "KP8_3_QB_DO" := "FB_KP8_DB_3".KP8.Rohdaten.QB_DO;

   //KP8_4
   "FB_KP8_DB_4"();
   "KP8_4_QB_Rot" := "FB_KP8_DB_4".KP8.Rohdaten.QB_Rot;
   "KP8_4_QB_Gruen" := "FB_KP8_DB_4".KP8.Rohdaten.QB_Gruen;
   "KP8_4_QB_Blau" := "FB_KP8_DB_4".KP8.Rohdaten.QB_Blau;
   "KP8_4_QB_DO" := "FB_KP8_DB_4".KP8.Rohdaten.QB_DO;

   //KP8_5
   "FB_KP8_DB_5"();
   "KP8_5_QB_Rot" := "FB_KP8_DB_5".KP8.Rohdaten.QB_Rot;
   "KP8_5_QB_Gruen" := "FB_KP8_DB_5".KP8.Rohdaten.QB_Gruen;
   "KP8_5_QB_Blau" := "FB_KP8_DB_5".KP8.Rohdaten.QB_Blau;
   "KP8_5_QB_DO" := "FB_KP8_DB_5".KP8.Rohdaten.QB_DO;

   //KP8_6
   "FB_KP8_DB_6"();
   "KP8_6_QB_Rot" := "FB_KP8_DB_6".KP8.Rohdaten.QB_Rot;
   "KP8_6_QB_Gruen" := "FB_KP8_DB_6".KP8.Rohdaten.QB_Gruen;
   "KP8_6_QB_Blau" := "FB_KP8_DB_6".KP8.Rohdaten.QB_Blau;
   "KP8_6_QB_DO" := "FB_KP8_DB_6".KP8.Rohdaten.QB_DO;

   //KP8_7
   "FB_KP8_DB_7"();
   "KP8_7_QB_Rot" := "FB_KP8_DB_7".KP8.Rohdaten.QB_Rot;
   "KP8_7_QB_Gruen" := "FB_KP8_DB_7".KP8.Rohdaten.QB_Gruen;
   "KP8_7_QB_Blau" := "FB_KP8_DB_7".KP8.Rohdaten.QB_Blau;
   "KP8_7_QB_DO" := "FB_KP8_DB_7".KP8.Rohdaten.QB_DO;

   //KP8_8
   "FB_KP8_DB_8"();
   "KP8_8_QB_Rot" := "FB_KP8_DB_8".KP8.Rohdaten.QB_Rot;
   "KP8_8_QB_Gruen" := "FB_KP8_DB_8".KP8.Rohdaten.QB_Gruen;
   "KP8_8_QB_Blau" := "FB_KP8_DB_8".KP8.Rohdaten.QB_Blau;
   "KP8_8_QB_DO" := "FB_KP8_DB_8".KP8.Rohdaten.QB_DO;

   //KP8_9
   "FB_KP8_DB_9"();
   "KP8_9_QB_Rot" := "FB_KP8_DB_9".KP8.Rohdaten.QB_Rot;
   "KP8_9_QB_Gruen" := "FB_KP8_DB_9".KP8.Rohdaten.QB_Gruen;
   "KP8_9_QB_Blau" := "FB_KP8_DB_9".KP8.Rohdaten.QB_Blau;
   "KP8_9_QB_DO" := "FB_KP8_DB_9".KP8.Rohdaten.QB_DO;

   //KP8_10
   "FB_KP8_DB_10"();
   "KP8_10_QB_Rot" := "FB_KP8_DB_10".KP8.Rohdaten.QB_Rot;
   "KP8_10_QB_Gruen" := "FB_KP8_DB_10".KP8.Rohdaten.QB_Gruen;
   "KP8_10_QB_Blau" := "FB_KP8_DB_10".KP8.Rohdaten.QB_Blau;
   "KP8_10_QB_DO" := "FB_KP8_DB_10".KP8.Rohdaten.QB_DO;

   //KP8_11
   "FB_KP8_DB_11"();
   "KP8_11_QB_Rot" := "FB_KP8_DB_11".KP8.Rohdaten.QB_Rot;
   "KP8_11_QB_Gruen" := "FB_KP8_DB_11".KP8.Rohdaten.QB_Gruen;
   "KP8_11_QB_Blau" := "FB_KP8_DB_11".KP8.Rohdaten.QB_Blau;
   "KP8_11_QB_DO" := "FB_KP8_DB_11".KP8.Rohdaten.QB_DO;

   //KP8_12
   "FB_KP8_DB_12"();
   "KP8_12_QB_Rot" := "FB_KP8_DB_12".KP8.Rohdaten.QB_Rot;
   "KP8_12_QB_Gruen" := "FB_KP8_DB_12".KP8.Rohdaten.QB_Gruen;
   "KP8_12_QB_Blau" := "FB_KP8_DB_12".KP8.Rohdaten.QB_Blau;
   "KP8_12_QB_DO" := "FB_KP8_DB_12".KP8.Rohdaten.QB_DO;

   //KP8_13
   "FB_KP8_DB_13"();
   "KP8_13_QB_Rot" := "FB_KP8_DB_13".KP8.Rohdaten.QB_Rot;
   "KP8_13_QB_Gruen" := "FB_KP8_DB_13".KP8.Rohdaten.QB_Gruen;
   "KP8_13_QB_Blau" := "FB_KP8_DB_13".KP8.Rohdaten.QB_Blau;
   "KP8_13_QB_DO" := "FB_KP8_DB_13".KP8.Rohdaten.QB_DO;

   //KP8_14
   "FB_KP8_DB_14"();
   "KP8_14_QB_Rot" := "FB_KP8_DB_14".KP8.Rohdaten.QB_Rot;
   "KP8_14_QB_Gruen" := "FB_KP8_DB_14".KP8.Rohdaten.QB_Gruen;
   "KP8_14_QB_Blau" := "FB_KP8_DB_14".KP8.Rohdaten.QB_Blau;
   "KP8_14_QB_DO" := "FB_KP8_DB_14".KP8.Rohdaten.QB_DO;

   //KP8_15
   "FB_KP8_DB_15"();
   "KP8_15_QB_Rot" := "FB_KP8_DB_15".KP8.Rohdaten.QB_Rot;
   "KP8_15_QB_Gruen" := "FB_KP8_DB_15".KP8.Rohdaten.QB_Gruen;
   "KP8_15_QB_Blau" := "FB_KP8_DB_15".KP8.Rohdaten.QB_Blau;
   "KP8_15_QB_DO" := "FB_KP8_DB_15".KP8.Rohdaten.QB_DO;

   //KP8_16
   "FB_KP8_DB_16"();
   "KP8_16_QB_Rot" := "FB_KP8_DB_16".KP8.Rohdaten.QB_Rot;
   "KP8_16_QB_Gruen" := "FB_KP8_DB_16".KP8.Rohdaten.QB_Gruen;
   "KP8_16_QB_Blau" := "FB_KP8_DB_16".KP8.Rohdaten.QB_Blau;
   "KP8_16_QB_DO" := "FB_KP8_DB_16".KP8.Rohdaten.QB_DO;

   //KP8_17
   "FB_KP8_DB_17"();
   "KP8_17_QB_Rot" := "FB_KP8_DB_17".KP8.Rohdaten.QB_Rot;
   "KP8_17_QB_Gruen" := "FB_KP8_DB_17".KP8.Rohdaten.QB_Gruen;
   "KP8_17_QB_Blau" := "FB_KP8_DB_17".KP8.Rohdaten.QB_Blau;
   "KP8_17_QB_DO" := "FB_KP8_DB_17".KP8.Rohdaten.QB_DO;

   //KP8_18
   "FB_KP8_DB_18"();
   "KP8_18_QB_Rot" := "FB_KP8_DB_18".KP8.Rohdaten.QB_Rot;
   "KP8_18_QB_Gruen" := "FB_KP8_DB_18".KP8.Rohdaten.QB_Gruen;
   "KP8_18_QB_Blau" := "FB_KP8_DB_18".KP8.Rohdaten.QB_Blau;
   "KP8_18_QB_DO" := "FB_KP8_DB_18".KP8.Rohdaten.QB_DO;

   //KP8_19
   "FB_KP8_DB_19"();
   "KP8_19_QB_Rot" := "FB_KP8_DB_19".KP8.Rohdaten.QB_Rot;
   "KP8_19_QB_Gruen" := "FB_KP8_DB_19".KP8.Rohdaten.QB_Gruen;
   "KP8_19_QB_Blau" := "FB_KP8_DB_19".KP8.Rohdaten.QB_Blau;
   "KP8_19_QB_DO" := "FB_KP8_DB_19".KP8.Rohdaten.QB_DO;

   //KP8_20
   "FB_KP8_DB_20"();
   "KP8_20_QB_Rot" := "FB_KP8_DB_20".KP8.Rohdaten.QB_Rot;
   "KP8_20_QB_Gruen" := "FB_KP8_DB_20".KP8.Rohdaten.QB_Gruen;
   "KP8_20_QB_Blau" := "FB_KP8_DB_20".KP8.Rohdaten.QB_Blau;
   "KP8_20_QB_DO" := "FB_KP8_DB_20".KP8.Rohdaten.QB_DO;

   //KP8_21
   "FB_KP8_DB_21"();
   "KP8_21_QB_Rot" := "FB_KP8_DB_21".KP8.Rohdaten.QB_Rot;
   "KP8_21_QB_Gruen" := "FB_KP8_DB_21".KP8.Rohdaten.QB_Gruen;
   "KP8_21_QB_Blau" := "FB_KP8_DB_21".KP8.Rohdaten.QB_Blau;
   "KP8_21_QB_DO" := "FB_KP8_DB_21".KP8.Rohdaten.QB_DO;

   //KP8_22
   "FB_KP8_DB_22"();
   "KP8_22_QB_Rot" := "FB_KP8_DB_22".KP8.Rohdaten.QB_Rot;
   "KP8_22_QB_Gruen" := "FB_KP8_DB_22".KP8.Rohdaten.QB_Gruen;
   "KP8_22_QB_Blau" := "FB_KP8_DB_22".KP8.Rohdaten.QB_Blau;
   "KP8_22_QB_DO" := "FB_KP8_DB_22".KP8.Rohdaten.QB_DO;

   //KP8_23
   "FB_KP8_DB_23"();
   "KP8_23_QB_Rot" := "FB_KP8_DB_23".KP8.Rohdaten.QB_Rot;
   "KP8_23_QB_Gruen" := "FB_KP8_DB_23".KP8.Rohdaten.QB_Gruen;
   "KP8_23_QB_Blau" := "FB_KP8_DB_23".KP8.Rohdaten.QB_Blau;
   "KP8_23_QB_DO" := "FB_KP8_DB_23".KP8.Rohdaten.QB_DO;

   //KP8_24
   "FB_KP8_DB_24"();
   "KP8_24_QB_Rot" := "FB_KP8_DB_24".KP8.Rohdaten.QB_Rot;
   "KP8_24_QB_Gruen" := "FB_KP8_DB_24".KP8.Rohdaten.QB_Gruen;
   "KP8_24_QB_Blau" := "FB_KP8_DB_24".KP8.Rohdaten.QB_Blau;
   "KP8_24_QB_DO" := "FB_KP8_DB_24".KP8.Rohdaten.QB_DO;

   //KP8_25
   "FB_KP8_DB_25"();
   "KP8_25_QB_Rot" := "FB_KP8_DB_25".KP8.Rohdaten.QB_Rot;
   "KP8_25_QB_Gruen" := "FB_KP8_DB_25".KP8.Rohdaten.QB_Gruen;
   "KP8_25_QB_Blau" := "FB_KP8_DB_25".KP8.Rohdaten.QB_Blau;
   "KP8_25_QB_DO" := "FB_KP8_DB_25".KP8.Rohdaten.QB_DO;

   //KP8_26
   "FB_KP8_DB_26"();
   "KP8_26_QB_Rot" := "FB_KP8_DB_26".KP8.Rohdaten.QB_Rot;
   "KP8_26_QB_Gruen" := "FB_KP8_DB_26".KP8.Rohdaten.QB_Gruen;
   "KP8_26_QB_Blau" := "FB_KP8_DB_26".KP8.Rohdaten.QB_Blau;
   "KP8_26_QB_DO" := "FB_KP8_DB_26".KP8.Rohdaten.QB_DO;

   //KP8_27
   "FB_KP8_DB_27"();
   "KP8_27_QB_Rot" := "FB_KP8_DB_27".KP8.Rohdaten.QB_Rot;
   "KP8_27_QB_Gruen" := "FB_KP8_DB_27".KP8.Rohdaten.QB_Gruen;
   "KP8_27_QB_Blau" := "FB_KP8_DB_27".KP8.Rohdaten.QB_Blau;
   "KP8_27_QB_DO" := "FB_KP8_DB_27".KP8.Rohdaten.QB_DO;

   //KP8_28
   "FB_KP8_DB_28"();
   "KP8_28_QB_Rot" := "FB_KP8_DB_28".KP8.Rohdaten.QB_Rot;
   "KP8_28_QB_Gruen" := "FB_KP8_DB_28".KP8.Rohdaten.QB_Gruen;
   "KP8_28_QB_Blau" := "FB_KP8_DB_28".KP8.Rohdaten.QB_Blau;
   "KP8_28_QB_DO" := "FB_KP8_DB_28".KP8.Rohdaten.QB_DO;
END_REGION

REGION Network 5 (SCL): Fehlermeldungen
   "FC_Fehlermeldungen"();
END_REGION

REGION Network 6 (SCL): Not-Halt
   "FC_Not_Halt"(NOT "Not-Aus ist OK");
END_REGION

REGION Network 7 (SCL): Not-Aus Reset
       "Not-Aus Reset" := "DB_IPC_to_CPU".Not_Halt_Reset;     // %Q4.7
END_REGION
END_ORGANIZATION_BLOCK

FUNCTION_BLOCK "FB_Ansteuerung_KP8"   // FB5, SCL
{ S7_Optimized_Access := 'TRUE' }
VERSION : 0.1
// stored: AutoNumber true, IsIECCheckEnabled false, IsRetainMemResEnabled false, MemoryReserve 100, SetENOAutomatically false, UDAEnableTagReadback false
   VAR
      KP8 { ExternalAccessible := 'False'; ExternalVisible := 'False'; ExternalWritable := 'False'} : "UDT_KP8";
   END_VAR
   VAR_TEMP
      i : USInt;
      Maske : Byte;
   END_VAR
BEGIN
   // 1) Eingänge dekodieren
   FOR #i := 0 TO 7 DO
       #Maske := SHL(IN := BYTE#1, N := #i);

       #KP8.Taste[#i] := (#KP8.Rohdaten.IB_Tasten AND #Maske) <> BYTE#0;
       #KP8.DI[#i] := (#KP8.Rohdaten.IB_DI AND #Maske) <> BYTE#0;
   END_FOR;

   // 2) Ausgänge neu aufbauen
   #KP8.Rohdaten.QB_Rot := BYTE#0;
   #KP8.Rohdaten.QB_Gruen := BYTE#0;
   #KP8.Rohdaten.QB_Blau := BYTE#0;
   #KP8.Rohdaten.QB_DO := BYTE#0;

   // 3) LEDs in Bytes umsetzen
   FOR #i := 0 TO 7 DO
       #Maske := SHL(IN := BYTE#1, N := #i);

       CASE #KP8.LED[#i] OF
           0: // Aus
               ;

           1: // Rot
               #KP8.Rohdaten.QB_Rot := #KP8.Rohdaten.QB_Rot OR #Maske;

           2: // Grün
               #KP8.Rohdaten.QB_Gruen := #KP8.Rohdaten.QB_Gruen OR #Maske;

           3: // Blau
               #KP8.Rohdaten.QB_Blau := #KP8.Rohdaten.QB_Blau OR #Maske;

           4: // Gelb
               #KP8.Rohdaten.QB_Rot := #KP8.Rohdaten.QB_Rot OR #Maske;
               #KP8.Rohdaten.QB_Gruen := #KP8.Rohdaten.QB_Gruen OR #Maske;

           5: // Weiß
               #KP8.Rohdaten.QB_Rot := #KP8.Rohdaten.QB_Rot OR #Maske;
               #KP8.Rohdaten.QB_Gruen := #KP8.Rohdaten.QB_Gruen OR #Maske;
               #KP8.Rohdaten.QB_Blau := #KP8.Rohdaten.QB_Blau OR #Maske;
       END_CASE;
   END_FOR;

   // 4) Digitale Ausgänge umsetzen
   FOR #i := 0 TO 7 DO
       #Maske := SHL(IN := BYTE#1, N := #i);

       IF #KP8.DO[#i] THEN
           #KP8.Rohdaten.QB_DO := #KP8.Rohdaten.QB_DO OR #Maske;
       END_IF;
   END_FOR;
END_FUNCTION_BLOCK

FUNCTION_BLOCK "FB_Anlagensteuerung"   // FB9, SCL
{ S7_Optimized_Access := 'TRUE' }
VERSION : 0.9
// stored: AutoNumber true, IsIECCheckEnabled false, IsRetainMemResEnabled false, MemoryReserve 100, SetENOAutomatically false, UDAEnableTagReadback false
   VAR_INPUT
      Blink_Takt : Bool;
      Clock_10Hz : Bool;
      Not_Halt_Aktiv : Bool;
   END_VAR
   VAR
      Auftragsmanager { S7_SetPoint := 'True'} : "FB_Auftragsmanager";
      Bad { S7_SetPoint := 'True'} : Array[1.."c_Anzahl_Bad"] of "FB_Bad";
      Heizung { S7_SetPoint := 'True'} : "FB_Heizungssteuerung";
      Blink_Zaehler : Int;
      M_10Hz_Alt : Bool;
   END_VAR
   VAR_TEMP
      "b" : Int;
      lampentest : Bool;
   END_VAR
BEGIN

       IF #Clock_10Hz AND NOT #M_10Hz_Alt THEN #Blink_Zaehler:=#Blink_Zaehler+1; IF #Blink_Zaehler>19 THEN #Blink_Zaehler:=0; END_IF; END_IF;
       #M_10Hz_Alt:=#Clock_10Hz;
       #lampentest:="DB_IPC_to_CPU".Lampentest;


       "FC_IO_Mapping"(Richtung:=1);
       #Auftragsmanager(Auftraege:="DB_IPC_to_CPU".Auftrag, Bad_Konfig:="DB_Bad_Konfig".Bad_Konfig);
       FOR #b:=1 TO "c_Anzahl_Bad" DO
           #Bad[#b](Blink_Takt:=#Blink_Takt, Lampentest:=#lampentest, Blink_Zaehler:=#Blink_Zaehler,
                    Not_Halt_Aktiv:=#Not_Halt_Aktiv, Zustand:="DB_IPC_to_CPU".Zustand[#b], BadNr:=#b,
                    Bad_Konfig:="DB_Bad_Konfig".Bad_Konfig[#b],
                    Auftraege:="DB_IPC_to_CPU".Auftrag,
                    Handbetrieb:="DB_IPC_to_CPU".Handbetrieb[#b],
                    Leerlauf:="DB_IPC_to_CPU".Leerlauf[#b],
                    Standby:="DB_IPC_to_CPU".Standby[#b]);
       END_FOR;
       #Heizung();
       "FC_IO_Mapping"(Richtung:=2);
       "FC_KP8_Override"(Lampentest:=#lampentest, Blink_Takt:=#Blink_Takt);
       "FC_Rueckmeldung"(Not_Halt_Aktiv:=#Not_Halt_Aktiv);
END_FUNCTION_BLOCK

FUNCTION_BLOCK "FB_Auftragsmanager"   // FB8, SCL
{ S7_Optimized_Access := 'TRUE' }
VERSION : 0.4
// stored: AutoNumber true, IsIECCheckEnabled false, IsRetainMemResEnabled false, MemoryReserve 100, SetENOAutomatically false, UDAEnableTagReadback false
   VAR_IN_OUT
      Auftraege : Array[0..9] of "UDT_Prozessroute";
      Bad_Konfig : Array[1.."c_Anzahl_Bad"] of "UDT_Bad_Konfig";
   END_VAR
   VAR
      Freigabe_Alt : Array[0..9] of Bool;
   END_VAR
   VAR_TEMP
      i : Int;
      "b" : Int;
      w : Int;
      ersterBad : Int;
      naechsterBad : Int;
      aktSchrittIdx : Int;
      flanke_Freigabe : Bool;
      auftrag_laeuft : Bool;
      freier_platz : Int;
   END_VAR
BEGIN

       FOR #b:=1 TO "c_Anzahl_Bad" DO FOR #w:=1 TO 3 DO
           IF #Bad_Konfig[#b].WT[#w].WT_Entnommen THEN
               #i:=#Bad_Konfig[#b].WT[#w].Auftragsindex; #aktSchrittIdx:=#Bad_Konfig[#b].WT[#w].SchrittIndex;
               IF (#i>=0)AND(#i<=9) THEN
                   IF (#aktSchrittIdx+1)<#Auftraege[#i].Anzahl_Schritte THEN
                       // Naechster Schritt: erst pruefen ob Platz frei
                       #naechsterBad:=#Auftraege[#i].Schritte[#aktSchrittIdx+1].BadNr;
                       #freier_platz:=0;
                       IF (#naechsterBad>=1)AND(#naechsterBad<="c_Anzahl_Bad") THEN
                           IF #Bad_Konfig[#naechsterBad].Ausstattung.HatGleichrichter
                              AND (#Bad_Konfig[#naechsterBad].WT[1].Belegt OR #Bad_Konfig[#naechsterBad].WT[2].Belegt OR #Bad_Konfig[#naechsterBad].WT[3].Belegt) THEN
                               #freier_platz:=0;
                           ELSIF NOT #Bad_Konfig[#naechsterBad].WT[1].Belegt THEN #freier_platz:=1;
                           ELSIF NOT #Bad_Konfig[#naechsterBad].WT[2].Belegt THEN #freier_platz:=2;
                           ELSIF NOT #Bad_Konfig[#naechsterBad].WT[3].Belegt THEN #freier_platz:=3; END_IF;
                       END_IF;
                       IF #freier_platz>0 THEN
                           // Platz frei: altes Bad raeumen, neues Bad belegen
                           #Bad_Konfig[#b].WT[#w].Belegt:=FALSE; #Bad_Konfig[#b].WT[#w].Auftragsindex:=-1; #Bad_Konfig[#b].WT[#w].SchrittIndex:=-1;
                           #Bad_Konfig[#b].WT[#w].WT_Eingesetzt:=FALSE; #Bad_Konfig[#b].WT[#w].WT_Entnommen:=FALSE;
                           #Bad_Konfig[#b].WT[#w].Istzeit:=T#0s; #Bad_Konfig[#b].WT[#w].Restzeit:=T#0s;
                           #Bad_Konfig[#b].WT[#w].Zeit_Abgelaufen:=FALSE; #Bad_Konfig[#b].WT[#w].Krit_Zeit_Abgelaufen:=FALSE; #Bad_Konfig[#b].WT[#w].Vorwarn_Erreicht:=FALSE;
                           #Bad_Konfig[#naechsterBad].WT[#freier_platz].Auftragsindex:=#i; #Bad_Konfig[#naechsterBad].WT[#freier_platz].SchrittIndex:=#aktSchrittIdx+1;
                           #Bad_Konfig[#naechsterBad].WT[#freier_platz].Belegt:=TRUE; #Bad_Konfig[#naechsterBad].WT[#freier_platz].WT_Eingesetzt:=FALSE;
                           #Bad_Konfig[#naechsterBad].WT[#freier_platz].WT_Entnommen:=FALSE; #Bad_Konfig[#naechsterBad].WT[#freier_platz].Zeit_Abgelaufen:=FALSE;
                           #Bad_Konfig[#naechsterBad].WT[#freier_platz].Krit_Zeit_Abgelaufen:=FALSE; #Bad_Konfig[#naechsterBad].WT[#freier_platz].Vorwarn_Erreicht:=FALSE;
                           #Bad_Konfig[#naechsterBad].WT[#freier_platz].Protokoll_Neu:=FALSE;
                       END_IF;
                       // freier_platz=0: WT bleibt am alten Bad, naechsten Zyklus erneut pruefen
                   ELSE
                       // Letzter Schritt: raeumen und Auftrag abschliessen
                       #Bad_Konfig[#b].WT[#w].Belegt:=FALSE; #Bad_Konfig[#b].WT[#w].Auftragsindex:=-1; #Bad_Konfig[#b].WT[#w].SchrittIndex:=-1;
                       #Bad_Konfig[#b].WT[#w].WT_Eingesetzt:=FALSE; #Bad_Konfig[#b].WT[#w].WT_Entnommen:=FALSE;
                       #Bad_Konfig[#b].WT[#w].Istzeit:=T#0s; #Bad_Konfig[#b].WT[#w].Restzeit:=T#0s;
                       #Bad_Konfig[#b].WT[#w].Zeit_Abgelaufen:=FALSE; #Bad_Konfig[#b].WT[#w].Krit_Zeit_Abgelaufen:=FALSE; #Bad_Konfig[#b].WT[#w].Vorwarn_Erreicht:=FALSE;
                       #Auftraege[#i].Freigabe:=FALSE; #Freigabe_Alt[#i]:=FALSE;
                       "DB_CPU_to_IPC".Auftrag_Abgeschlossen[#i] := TRUE;
                   END_IF;
               END_IF;
           END_IF;
       END_FOR; END_FOR;
       FOR #i:=0 TO 9 DO IF #Auftraege[#i].Abbruch THEN
           FOR #b:=1 TO "c_Anzahl_Bad" DO FOR #w:=1 TO 3 DO
               IF #Bad_Konfig[#b].WT[#w].Auftragsindex=#i THEN
                   #Bad_Konfig[#b].WT[#w].Belegt:=FALSE; #Bad_Konfig[#b].WT[#w].Auftragsindex:=-1; #Bad_Konfig[#b].WT[#w].SchrittIndex:=-1;
                   #Bad_Konfig[#b].WT[#w].WT_Eingesetzt:=FALSE; #Bad_Konfig[#b].WT[#w].WT_Entnommen:=FALSE;
                   #Bad_Konfig[#b].WT[#w].Istzeit:=T#0s; #Bad_Konfig[#b].WT[#w].Restzeit:=T#0s;
                   #Bad_Konfig[#b].WT[#w].Zeit_Abgelaufen:=FALSE; #Bad_Konfig[#b].WT[#w].Krit_Zeit_Abgelaufen:=FALSE; #Bad_Konfig[#b].WT[#w].Vorwarn_Erreicht:=FALSE;
               END_IF;
           END_FOR; END_FOR;
           #Auftraege[#i].Freigabe:=FALSE; #Auftraege[#i].Abbruch:=FALSE; #Freigabe_Alt[#i]:=FALSE;
       END_IF; END_FOR;
       FOR #i:=0 TO 9 DO
           #flanke_Freigabe:=#Auftraege[#i].Freigabe AND NOT #Freigabe_Alt[#i]; #Freigabe_Alt[#i]:=#Auftraege[#i].Freigabe;
           // Auftrag_Abgeschlossen zuruecksetzen wenn IPC den Slot aufgeraeumt hat
           IF #Auftraege[#i].Anzahl_Schritte = 0 THEN "DB_CPU_to_IPC".Auftrag_Abgeschlossen[#i] := FALSE; END_IF;
           IF #Auftraege[#i].Freigabe AND NOT #Auftraege[#i].Abbruch THEN
               #auftrag_laeuft:=FALSE;
               FOR #b:=1 TO "c_Anzahl_Bad" DO FOR #w:=1 TO 3 DO IF #Bad_Konfig[#b].WT[#w].Auftragsindex=#i THEN #auftrag_laeuft:=TRUE; END_IF; END_FOR; END_FOR;
               IF NOT #auftrag_laeuft AND(#Auftraege[#i].Anzahl_Schritte>=1)AND(#Auftraege[#i].Anzahl_Schritte<=51) THEN
                   #ersterBad:=#Auftraege[#i].Schritte[0].BadNr;
                   IF (#ersterBad>=1)AND(#ersterBad<="c_Anzahl_Bad") THEN
                       #freier_platz:=0;
                       // Gleichrichter-Baeder: max. 1 WT gleichzeitig
                       IF #Bad_Konfig[#ersterBad].Ausstattung.HatGleichrichter
                          AND (#Bad_Konfig[#ersterBad].WT[1].Belegt OR #Bad_Konfig[#ersterBad].WT[2].Belegt OR #Bad_Konfig[#ersterBad].WT[3].Belegt) THEN
                           #freier_platz:=0;
                       ELSIF NOT #Bad_Konfig[#ersterBad].WT[1].Belegt THEN #freier_platz:=1;
                       ELSIF NOT #Bad_Konfig[#ersterBad].WT[2].Belegt THEN #freier_platz:=2;
                       ELSIF NOT #Bad_Konfig[#ersterBad].WT[3].Belegt THEN #freier_platz:=3; END_IF;
                       IF #freier_platz>0 THEN
                           #Bad_Konfig[#ersterBad].WT[#freier_platz].Auftragsindex:=#i; #Bad_Konfig[#ersterBad].WT[#freier_platz].SchrittIndex:=0;
                           #Bad_Konfig[#ersterBad].WT[#freier_platz].Belegt:=TRUE; #Bad_Konfig[#ersterBad].WT[#freier_platz].WT_Eingesetzt:=FALSE;
                           #Bad_Konfig[#ersterBad].WT[#freier_platz].WT_Entnommen:=FALSE; #Bad_Konfig[#ersterBad].WT[#freier_platz].Zeit_Abgelaufen:=FALSE;
                           #Bad_Konfig[#ersterBad].WT[#freier_platz].Krit_Zeit_Abgelaufen:=FALSE; #Bad_Konfig[#ersterBad].WT[#freier_platz].Vorwarn_Erreicht:=FALSE;
                           #Bad_Konfig[#ersterBad].WT[#freier_platz].Protokoll_Neu:=FALSE;
                       END_IF;
                   END_IF;
               END_IF;
           END_IF;
       END_FOR;
END_FUNCTION_BLOCK

FUNCTION_BLOCK "FB_Bad"   // FB7, SCL
{ S7_Optimized_Access := 'TRUE' }
VERSION : 0.9
// stored: AutoNumber true, IsIECCheckEnabled false, IsRetainMemResEnabled false, MemoryReserve 100, SetENOAutomatically false, UDAEnableTagReadback false
   VAR_INPUT
      Blink_Takt : Bool;
      Lampentest : Bool;
      Blink_Zaehler : Int;
      Not_Halt_Aktiv : Bool;
      Zustand : Int;   // 0=aus, 1=Leerlauf, 2=Standby
      BadNr : Int;
   END_VAR
   VAR_IN_OUT
      Bad_Konfig : "UDT_Bad_Konfig";
      Auftraege : Array[0..9] of "UDT_Prozessroute";
      Handbetrieb : "UDT_Handbetrieb";
      Leerlauf : "UDT_Peripherie_Soll";
      Standby : "UDT_Peripherie_Soll";
   END_VAR
   VAR
      Timer_WT { S7_SetPoint := 'True'} : Array[1..3] of TON_TIME;
      Timer_FU_Pause { S7_SetPoint := 'True'} : TON_TIME;
      Timer_FU_Pumpe_Stoerung { S7_SetPoint := 'True'} : TON_TIME;
      Timer_FU_WB1_Stoerung { S7_SetPoint := 'True'} : TON_TIME;
      Timer_FU_WB2_Stoerung { S7_SetPoint := 'True'} : TON_TIME;
      M_Ein_Any_Alt : Bool;
      M_Ent_Any_Alt : Bool;
   END_VAR
   VAR_TEMP
      w : Int;
      flanke_Ein : Bool;
      flanke_Ent : Bool;
      any_ein : Bool;
      any_ent : Bool;
      aktSchritt : "UDT_Badschritt";
      hat_Schritt : Bool;
      hw_ok : Bool;
      temp_ok : Bool;
      hw_ok_ohne_niveau : Bool;
      heiz1_ok : Bool;
      heiz2_ok : Bool;
      heiz_soll_max : Real;
      heiz_tol : Real;
      irgend_belegt : Bool;
      worst_ampel : Int;
      any_hupe : Bool;
      blink : Array[1..3] of Bool;
      pumpe_ein_any : Bool;
      us_ein_any : Bool;
      pumpe_fu_max : Real;
      irgend_eingesetzt : Bool;
      ent_prio_rest : Time;
      hand_aktiv : Bool;
      leerlauf_aktiv : Bool;
      standby_aktiv : Bool;
      irgend_aktiv : Bool;
      temp_abw : Real;
      aktZeit : DTL;
      retval : Int;
   END_VAR
BEGIN

       //== 1) Blinkmuster ==
       #blink[1] := (#Blink_Zaehler <= 9);
       #blink[2] := (#Blink_Zaehler <= 3) OR ((#Blink_Zaehler >= 8) AND (#Blink_Zaehler <= 11));
       #blink[3] := (#Blink_Zaehler <= 2) OR ((#Blink_Zaehler >= 6) AND (#Blink_Zaehler <= 8))
                   OR ((#Blink_Zaehler >= 12) AND (#Blink_Zaehler <= 14));

       //== 2) Ist-Werte ==
       #Bad_Konfig.Heizung_1_Ist := #Bad_Konfig.IO_Ein.Ist_Temperatur_1;
       #Bad_Konfig.Heizung_2_Ist := #Bad_Konfig.IO_Ein.Ist_Temperatur_2;

       //== 3) hw_ok ==
       #hw_ok := (#Bad_Konfig.IO_Ein.Niveau_OK      OR NOT #Bad_Konfig.Ausstattung.HatNiveau)
            AND (#Bad_Konfig.IO_Ein.Motorschutz_OK OR NOT #Bad_Konfig.Ausstattung.HatPumpe)
            AND (#Bad_Konfig.IO_Ein.FI_Schutz_OK   OR NOT (#Bad_Konfig.Ausstattung.HatHeizung_1 OR #Bad_Konfig.Ausstattung.HatHeizung_2))
            AND (#Bad_Konfig.IO_Ein.Kein_Uebertemp OR NOT (#Bad_Konfig.Ausstattung.HatHeizung_1 OR #Bad_Konfig.Ausstattung.HatHeizung_2))
            AND NOT #Not_Halt_Aktiv;

       // Pumpe darf auch ohne Niveau laufen (Niveau schuetzt nur die Heizung)
       #hw_ok_ohne_niveau :=
                (#Bad_Konfig.IO_Ein.Motorschutz_OK OR NOT #Bad_Konfig.Ausstattung.HatPumpe)
            AND (#Bad_Konfig.IO_Ein.FI_Schutz_OK   OR NOT (#Bad_Konfig.Ausstattung.HatHeizung_1 OR #Bad_Konfig.Ausstattung.HatHeizung_2))
            AND (#Bad_Konfig.IO_Ein.Kein_Uebertemp OR NOT (#Bad_Konfig.Ausstattung.HatHeizung_1 OR #Bad_Konfig.Ausstattung.HatHeizung_2))
            AND NOT #Not_Halt_Aktiv;

       //== 4) Belegung + Soll-Werte ==
       #irgend_belegt := FALSE;
       #pumpe_ein_any := FALSE; #us_ein_any := FALSE;
       #heiz_soll_max := 0.0; #heiz_tol := 5.0;
       #pumpe_fu_max := 0.0;

       FOR #w := 1 TO 3 DO
           IF #Bad_Konfig.WT[#w].Belegt THEN
               #irgend_belegt := TRUE;
               #hat_Schritt := (#Bad_Konfig.WT[#w].Auftragsindex >= 0) AND (#Bad_Konfig.WT[#w].Auftragsindex <= 9)
                          AND (#Bad_Konfig.WT[#w].SchrittIndex >= 0) AND (#Bad_Konfig.WT[#w].SchrittIndex <= 50);
               IF #hat_Schritt THEN
                   #aktSchritt := #Auftraege[#Bad_Konfig.WT[#w].Auftragsindex].Schritte[#Bad_Konfig.WT[#w].SchrittIndex];
                   IF #aktSchritt.Pumpe THEN #pumpe_ein_any := TRUE; END_IF;
                   IF #aktSchritt.Ultraschall THEN #us_ein_any := TRUE; END_IF;
                   IF #aktSchritt.Pumpe_FU_Soll > #pumpe_fu_max THEN #pumpe_fu_max := #aktSchritt.Pumpe_FU_Soll; END_IF;
                   IF #aktSchritt.Heizung > #heiz_soll_max THEN
                       #heiz_soll_max := #aktSchritt.Heizung;
                       #heiz_tol := #aktSchritt.Heizung_Toleranz;
                   END_IF;
               END_IF;
           END_IF;
       END_FOR;

       //== 5) Betriebsmodi ==
       #hand_aktiv := #Handbetrieb.Hand_Aktiv AND NOT #irgend_belegt AND NOT #Not_Halt_Aktiv;
       #Bad_Konfig.Hand_Aktiv_Intern := #hand_aktiv;
       #leerlauf_aktiv := (#Zustand = 1) AND NOT #irgend_belegt AND NOT #hand_aktiv
                         AND NOT #Not_Halt_Aktiv;
       #standby_aktiv := (#Zustand = 2) AND NOT #irgend_belegt AND NOT #hand_aktiv
                        AND NOT #Not_Halt_Aktiv;
       #irgend_aktiv := #irgend_belegt OR #hand_aktiv OR #leerlauf_aktiv OR #standby_aktiv;

       // Pruefen ob mindestens 1 WT eingesetzt ist
       #irgend_eingesetzt := FALSE;
       FOR #w := 1 TO 3 DO
           IF #Bad_Konfig.WT[#w].Belegt AND #Bad_Konfig.WT[#w].WT_Eingesetzt THEN #irgend_eingesetzt := TRUE; END_IF;
       END_FOR;

       IF #irgend_belegt THEN
           // Automatik: Heizung SOFORT bei Belegung (Vorheizen)
           IF #Bad_Konfig.Ausstattung.HatHeizung_1 THEN #Bad_Konfig.Heizung_1_Soll := #heiz_soll_max; END_IF;
           IF #Bad_Konfig.Ausstattung.HatHeizung_2 THEN #Bad_Konfig.Heizung_2_Soll := #heiz_soll_max; END_IF;
           // FU-Pause: 10s Ausrollzeit nach Auftragsstart (Uebergang Leerlauf->Automatik)
           #Timer_FU_Pause(IN := TRUE, PT := T#10s);
           // Alles andere ERST wenn mindestens 1 WT eingesetzt
           IF #irgend_eingesetzt THEN
               IF #Bad_Konfig.Ausstattung.HatPumpe THEN #Bad_Konfig.Pumpe_Ein := #pumpe_ein_any; END_IF;
               // Pumpe FU erst nach Ablauf der 10s Pause
               IF #Bad_Konfig.Ausstattung.HatPumpe_FU AND #Timer_FU_Pause.Q THEN
                   #Bad_Konfig.Pumpe_FU_Soll := #pumpe_fu_max;
               ELSIF #Bad_Konfig.Ausstattung.HatPumpe_FU THEN
                   #Bad_Konfig.Pumpe_FU_Soll := 0.0;
               END_IF;
               IF #Bad_Konfig.Ausstattung.HatUltraschall THEN #Bad_Konfig.Ultraschall_Ein := #us_ein_any; END_IF;
               IF #Bad_Konfig.Ausstattung.HatGleichrichter THEN
                   #Bad_Konfig.GR_Aktiv := #aktSchritt.GR_Aktiv;
                   #Bad_Konfig.GR_Strom_Soll := #aktSchritt.GR_Strom_Soll;
                   #Bad_Konfig.GR_Spannung_Soll := #aktSchritt.GR_Spannung_Soll;
                   #Bad_Konfig.GR_Pulsfrequenz := #aktSchritt.GR_Pulsfrequenz;
                   #Bad_Konfig.GR_DutyCycle := #aktSchritt.GR_DutyCycle;
               END_IF;
               IF #Bad_Konfig.Ausstattung.HatWarenbewegung_X AND #Timer_FU_Pause.Q THEN
                   #Bad_Konfig.Warenbewegung_X_Soll := #aktSchritt.Warenbewegung_X;
               ELSIF #Bad_Konfig.Ausstattung.HatWarenbewegung_X THEN
                   #Bad_Konfig.Warenbewegung_X_Soll := 0.0;
               END_IF;
               IF #Bad_Konfig.Ausstattung.HatWarenbewegung_Y AND #Timer_FU_Pause.Q THEN
                   #Bad_Konfig.Warenbewegung_Y_Soll := #aktSchritt.Warenbewegung_Y;
               ELSIF #Bad_Konfig.Ausstattung.HatWarenbewegung_Y THEN
                   #Bad_Konfig.Warenbewegung_Y_Soll := 0.0;
               END_IF;
           ELSE
               // Belegt aber kein WT eingesetzt: Aggregate aus
               #Bad_Konfig.Pumpe_Ein := FALSE;
               #Bad_Konfig.Pumpe_FU_Soll := 0.0;
               #Bad_Konfig.Ultraschall_Ein := FALSE;
               #Bad_Konfig.GR_Aktiv := FALSE;
               #Bad_Konfig.GR_Strom_Soll := 0.0; #Bad_Konfig.GR_Spannung_Soll := 0.0;
               #Bad_Konfig.GR_Pulsfrequenz := 0.0; #Bad_Konfig.GR_DutyCycle := 0.0;
           END_IF;
           // FU-Resets im Automatik immer FALSE
           #Bad_Konfig.WB1_Reset := FALSE;
           #Bad_Konfig.WB2_Reset := FALSE;
           #Bad_Konfig.IO_Aus.Pumpe_FU_Reset := FALSE;
       ELSIF #hand_aktiv THEN
           // Handbetrieb
           #Timer_FU_Pause(IN := FALSE, PT := T#10s);
           IF #Bad_Konfig.Ausstattung.HatHeizung_1 THEN #Bad_Konfig.Heizung_1_Soll := #Handbetrieb.Heizung_Soll; END_IF;
           IF #Bad_Konfig.Ausstattung.HatHeizung_2 THEN #Bad_Konfig.Heizung_2_Soll := #Handbetrieb.Heizung_Soll; END_IF;
           IF #Bad_Konfig.Ausstattung.HatPumpe THEN #Bad_Konfig.Pumpe_Ein := #Handbetrieb.Pumpe; END_IF;
           IF #Bad_Konfig.Ausstattung.HatPumpe_FU THEN #Bad_Konfig.Pumpe_FU_Soll := #Handbetrieb.Pumpe_FU_Soll; END_IF;
           IF #Bad_Konfig.Ausstattung.HatUltraschall THEN #Bad_Konfig.Ultraschall_Ein := #Handbetrieb.Ultraschall; END_IF;
           IF #Bad_Konfig.Ausstattung.HatGleichrichter THEN
               #Bad_Konfig.GR_Aktiv := #Handbetrieb.GR_Aktiv;
               #Bad_Konfig.GR_Strom_Soll := #Handbetrieb.GR_Strom_Soll;
               #Bad_Konfig.GR_Spannung_Soll := #Handbetrieb.GR_Spannung_Soll;
               #Bad_Konfig.GR_Pulsfrequenz := #Handbetrieb.GR_Pulsfrequenz;
               #Bad_Konfig.GR_DutyCycle := #Handbetrieb.GR_DutyCycle;
           END_IF;
           IF #Bad_Konfig.Ausstattung.HatWarenbewegung_X THEN #Bad_Konfig.Warenbewegung_X_Soll := #Handbetrieb.Warenbewegung_X; END_IF;
           IF #Bad_Konfig.Ausstattung.HatWarenbewegung_Y THEN #Bad_Konfig.Warenbewegung_Y_Soll := #Handbetrieb.Warenbewegung_Y; END_IF;
           #heiz_soll_max := #Handbetrieb.Heizung_Soll;
           // FU-Resets vom IPC durchreichen
           #Bad_Konfig.WB1_Reset := #Handbetrieb.WB1_Reset;
           #Bad_Konfig.WB2_Reset := #Handbetrieb.WB2_Reset;
           #Bad_Konfig.IO_Aus.Pumpe_FU_Reset := #Handbetrieb.Pumpe_FU_Reset;
       ELSIF #leerlauf_aktiv THEN
           // Leerlauf (Zustand 1): Bad betriebsbereit halten
           #Timer_FU_Pause(IN := FALSE, PT := T#10s);
           IF #Bad_Konfig.Ausstattung.HatHeizung_1 THEN #Bad_Konfig.Heizung_1_Soll := #Leerlauf.Heizung_Soll; END_IF;
           IF #Bad_Konfig.Ausstattung.HatHeizung_2 THEN #Bad_Konfig.Heizung_2_Soll := #Leerlauf.Heizung_Soll; END_IF;
           IF #Bad_Konfig.Ausstattung.HatPumpe THEN #Bad_Konfig.Pumpe_Ein := #Leerlauf.Pumpe; END_IF;
           IF #Bad_Konfig.Ausstattung.HatPumpe_FU THEN #Bad_Konfig.Pumpe_FU_Soll := #Leerlauf.Pumpe_FU_Soll; END_IF;
           IF #Bad_Konfig.Ausstattung.HatUltraschall THEN #Bad_Konfig.Ultraschall_Ein := #Leerlauf.Ultraschall; END_IF;
           IF #Bad_Konfig.Ausstattung.HatWarenbewegung_X THEN #Bad_Konfig.Warenbewegung_X_Soll := #Leerlauf.Warenbewegung_X; END_IF;
           IF #Bad_Konfig.Ausstattung.HatWarenbewegung_Y THEN #Bad_Konfig.Warenbewegung_Y_Soll := #Leerlauf.Warenbewegung_Y; END_IF;
           IF #Bad_Konfig.Ausstattung.HatGleichrichter THEN
               #Bad_Konfig.GR_Aktiv := #Leerlauf.GR_Aktiv;
               #Bad_Konfig.GR_Strom_Soll := #Leerlauf.GR_Strom_Soll;
               #Bad_Konfig.GR_Spannung_Soll := #Leerlauf.GR_Spannung_Soll;
           END_IF;
           #heiz_soll_max := #Leerlauf.Heizung_Soll;
           #Bad_Konfig.WB1_Reset := FALSE; #Bad_Konfig.WB2_Reset := FALSE;
           #Bad_Konfig.IO_Aus.Pumpe_FU_Reset := FALSE;
       ELSIF (#Zustand = 2) AND NOT #irgend_belegt AND NOT #hand_aktiv AND NOT #Not_Halt_Aktiv THEN
           // Standby (Zustand 2): Abgesenkte Temperatur, Aggregate pro Bad konfigurierbar
           #Timer_FU_Pause(IN := FALSE, PT := T#10s);
           IF #Bad_Konfig.Ausstattung.HatHeizung_1 THEN #Bad_Konfig.Heizung_1_Soll := #Standby.Heizung_Soll; END_IF;
           IF #Bad_Konfig.Ausstattung.HatHeizung_2 THEN #Bad_Konfig.Heizung_2_Soll := #Standby.Heizung_Soll; END_IF;
           IF #Bad_Konfig.Ausstattung.HatPumpe THEN #Bad_Konfig.Pumpe_Ein := #Standby.Pumpe; END_IF;
           IF #Bad_Konfig.Ausstattung.HatPumpe_FU THEN #Bad_Konfig.Pumpe_FU_Soll := #Standby.Pumpe_FU_Soll; END_IF;
           IF #Bad_Konfig.Ausstattung.HatUltraschall THEN #Bad_Konfig.Ultraschall_Ein := #Standby.Ultraschall; END_IF;
           IF #Bad_Konfig.Ausstattung.HatWarenbewegung_X THEN #Bad_Konfig.Warenbewegung_X_Soll := #Standby.Warenbewegung_X; END_IF;
           IF #Bad_Konfig.Ausstattung.HatWarenbewegung_Y THEN #Bad_Konfig.Warenbewegung_Y_Soll := #Standby.Warenbewegung_Y; END_IF;
           IF #Bad_Konfig.Ausstattung.HatGleichrichter THEN
               #Bad_Konfig.GR_Aktiv := #Standby.GR_Aktiv;
               #Bad_Konfig.GR_Strom_Soll := #Standby.GR_Strom_Soll;
               #Bad_Konfig.GR_Spannung_Soll := #Standby.GR_Spannung_Soll;
           END_IF;
           #heiz_soll_max := #Standby.Heizung_Soll;
           #Bad_Konfig.WB1_Reset := FALSE; #Bad_Konfig.WB2_Reset := FALSE;
           #Bad_Konfig.IO_Aus.Pumpe_FU_Reset := FALSE;
       ELSE
           // Zustand 0 oder undefiniert: alles aus
           #Timer_FU_Pause(IN := FALSE, PT := T#10s);
           #Bad_Konfig.Heizung_1_Soll := 0.0;
           #Bad_Konfig.Heizung_2_Soll := 0.0;
           #Bad_Konfig.Pumpe_Ein := FALSE;
           #Bad_Konfig.Pumpe_FU_Soll := 0.0;
           #Bad_Konfig.Ultraschall_Ein := FALSE;
           #Bad_Konfig.Warenbewegung_X_Soll := 0.0;
           #Bad_Konfig.Warenbewegung_Y_Soll := 0.0;
           #Bad_Konfig.GR_Aktiv := FALSE;
           #Bad_Konfig.GR_Strom_Soll := 0.0; #Bad_Konfig.GR_Spannung_Soll := 0.0;
           #Bad_Konfig.GR_Pulsfrequenz := 0.0; #Bad_Konfig.GR_DutyCycle := 0.0;
           #Bad_Konfig.WB1_Reset := FALSE; #Bad_Konfig.WB2_Reset := FALSE;
           #Bad_Konfig.IO_Aus.Pumpe_FU_Reset := FALSE;
       END_IF;

       //== 6) temp_ok ==
       #heiz1_ok := TRUE; #heiz2_ok := TRUE;
       IF #heiz_soll_max > 0.0 AND #irgend_aktiv THEN
           IF #heiz_tol <= 0.0 THEN #heiz_tol := 5.0; END_IF;
           IF #Bad_Konfig.Ausstattung.HatHeizung_1 THEN
               #heiz1_ok := ABS(#Bad_Konfig.IO_Ein.Ist_Temperatur_1 - #heiz_soll_max) <= #heiz_tol;
           END_IF;
           IF #Bad_Konfig.Ausstattung.HatHeizung_2 THEN
               #heiz2_ok := ABS(#Bad_Konfig.IO_Ein.Ist_Temperatur_2 - #heiz_soll_max) <= #heiz_tol;
           END_IF;
       END_IF;
       #temp_ok := #heiz1_ok AND #heiz2_ok;
       #Bad_Konfig.Betriebsbereit := #hw_ok AND #temp_ok;

       //== 7) Flanke ==
       #any_ein := #Bad_Konfig.IO_Ein.WT_Einsetzen[1] OR #Bad_Konfig.IO_Ein.WT_Einsetzen[2] OR #Bad_Konfig.IO_Ein.WT_Einsetzen[3];
       #any_ent := #Bad_Konfig.IO_Ein.WT_Entnehmen[1] OR #Bad_Konfig.IO_Ein.WT_Entnehmen[2] OR #Bad_Konfig.IO_Ein.WT_Entnehmen[3];
       #flanke_Ein := #any_ein AND NOT #M_Ein_Any_Alt;
       #flanke_Ent := #any_ent AND NOT #M_Ent_Any_Alt;
       #M_Ein_Any_Alt := #any_ein;
       #M_Ent_Any_Alt := #any_ent;

       //== 8) Pro-WT Ablauf ==
       FOR #w := 1 TO 3 DO
           #hat_Schritt := #Bad_Konfig.WT[#w].Belegt
               AND (#Bad_Konfig.WT[#w].Auftragsindex >= 0) AND (#Bad_Konfig.WT[#w].Auftragsindex <= 9)
               AND (#Bad_Konfig.WT[#w].SchrittIndex >= 0) AND (#Bad_Konfig.WT[#w].SchrittIndex <= 50);
           IF #hat_Schritt THEN
               #aktSchritt := #Auftraege[#Bad_Konfig.WT[#w].Auftragsindex].Schritte[#Bad_Konfig.WT[#w].SchrittIndex];
               IF NOT #Bad_Konfig.WT[#w].WT_Eingesetzt THEN
                   IF #flanke_Ein AND #Bad_Konfig.IO_Ein.WT_Einsetzen[#w] AND #hw_ok AND #temp_ok THEN
                       #Bad_Konfig.WT[#w].WT_Eingesetzt := TRUE;
                       #Bad_Konfig.WT[#w].WT_Entnommen := FALSE;
                       #Bad_Konfig.WT[#w].Istzeit := T#0s;
                       #Bad_Konfig.WT[#w].Zeit_Abgelaufen := FALSE;
                       #Bad_Konfig.WT[#w].Krit_Zeit_Abgelaufen := FALSE;
                       #Bad_Konfig.WT[#w].Vorwarn_Erreicht := FALSE;
                       #Bad_Konfig.WT[#w].Stoerung_Aufgetreten := FALSE;
                       #Bad_Konfig.WT[#w].Temp_Abweichung_Max := 0.0;
                       #Bad_Konfig.WT[#w].Temp_Toleranz_Eingehalten := TRUE;
                       #Bad_Konfig.WT[#w].Zeitueberschreitung := T#0s;
                       #Bad_Konfig.WT[#w].Protokoll_Neu := FALSE;
                       #retval := RD_LOC_T(OUT => #aktZeit);
                       #Bad_Konfig.WT[#w].Zeitstempel_Eingesetzt := #aktZeit;
                   END_IF;
               ELSE
                   #Timer_WT[#w](IN := TRUE, PT := T#24h);
                   #Bad_Konfig.WT[#w].Istzeit := #Timer_WT[#w].ET;
                   IF #Timer_WT[#w].ET < #aktSchritt.Verweilzeit THEN
                       #Bad_Konfig.WT[#w].Restzeit := #aktSchritt.Verweilzeit - #Timer_WT[#w].ET;
                   ELSE #Bad_Konfig.WT[#w].Restzeit := T#0s; END_IF;
                   IF #Timer_WT[#w].ET >= (#aktSchritt.Verweilzeit - #aktSchritt.Vorwarnzeit) THEN #Bad_Konfig.WT[#w].Vorwarn_Erreicht := TRUE; END_IF;
                   IF #Timer_WT[#w].ET >= #aktSchritt.Verweilzeit THEN #Bad_Konfig.WT[#w].Zeit_Abgelaufen := TRUE; END_IF;
                   IF #Timer_WT[#w].ET >= #aktSchritt.Kritische_Zeit THEN #Bad_Konfig.WT[#w].Krit_Zeit_Abgelaufen := TRUE; END_IF;
                   IF NOT #hw_ok THEN #Bad_Konfig.WT[#w].Stoerung_Aufgetreten := TRUE; END_IF;
                   IF #Bad_Konfig.Ausstattung.HatHeizung_1 AND (#aktSchritt.Heizung > 0.0) THEN
                       #temp_abw := ABS(#Bad_Konfig.IO_Ein.Ist_Temperatur_1 - #aktSchritt.Heizung);
                       IF #temp_abw > #Bad_Konfig.WT[#w].Temp_Abweichung_Max THEN #Bad_Konfig.WT[#w].Temp_Abweichung_Max := #temp_abw; END_IF;
                       IF #temp_abw > #aktSchritt.Heizung_Toleranz THEN #Bad_Konfig.WT[#w].Temp_Toleranz_Eingehalten := FALSE; END_IF;
                   END_IF;
                   IF #flanke_Ent AND #Bad_Konfig.IO_Ein.WT_Entnehmen[#w] THEN
                       #Bad_Konfig.WT[#w].WT_Entnommen := TRUE;
                       #Timer_WT[#w](IN := FALSE, PT := T#0s);
                       IF #Bad_Konfig.WT[#w].Istzeit > #aktSchritt.Verweilzeit THEN
                           #Bad_Konfig.WT[#w].Zeitueberschreitung := #Bad_Konfig.WT[#w].Istzeit - #aktSchritt.Verweilzeit;
                       ELSE #Bad_Konfig.WT[#w].Zeitueberschreitung := T#0s; END_IF;
                       #retval := RD_LOC_T(OUT => #aktZeit);
                       #Bad_Konfig.WT[#w].Zeitstempel_Entnommen := #aktZeit;
                       #Bad_Konfig.WT[#w].Protokoll_Neu := TRUE;
                   END_IF;
               END_IF;
           ELSE
               #Timer_WT[#w](IN := FALSE, PT := T#0s);
               #Bad_Konfig.WT[#w].Istzeit := T#0s; #Bad_Konfig.WT[#w].Restzeit := T#0s;
               #Bad_Konfig.WT[#w].Zeit_Abgelaufen := FALSE;
               #Bad_Konfig.WT[#w].Krit_Zeit_Abgelaufen := FALSE;
               #Bad_Konfig.WT[#w].Vorwarn_Erreicht := FALSE;
           END_IF;
       END_FOR;

       //== 9) Ampel ==
       #worst_ampel := 0; #any_hupe := FALSE;
       IF #Not_Halt_Aktiv THEN
           // Not-Halt: ALLE Ampeln rot blinken, unabhaengig von Belegung
           #worst_ampel := 4;  // rot blink (nicht konstant, damit man sieht: Not-Halt, nicht HW-Stoerung)
       ELSIF NOT #hw_ok AND #irgend_aktiv THEN
           #worst_ampel := 6;  // rot konstant = HW-Stoerung
       ELSIF #hand_aktiv AND NOT #irgend_belegt THEN
           #worst_ampel := 2;
       ELSE
           FOR #w := 1 TO 3 DO
               #hat_Schritt := #Bad_Konfig.WT[#w].Belegt
                   AND (#Bad_Konfig.WT[#w].Auftragsindex >= 0) AND (#Bad_Konfig.WT[#w].Auftragsindex <= 9)
                   AND (#Bad_Konfig.WT[#w].SchrittIndex >= 0) AND (#Bad_Konfig.WT[#w].SchrittIndex <= 50);
               IF #hat_Schritt THEN
                   IF #Bad_Konfig.WT[#w].WT_Eingesetzt THEN
                       #aktSchritt := #Auftraege[#Bad_Konfig.WT[#w].Auftragsindex].Schritte[#Bad_Konfig.WT[#w].SchrittIndex];
                       IF #Bad_Konfig.WT[#w].Krit_Zeit_Abgelaufen AND #aktSchritt.Alarm_Aktiv THEN
                           IF 5 > #worst_ampel THEN #worst_ampel := 5; END_IF; #any_hupe := TRUE;
                       ELSIF #Bad_Konfig.WT[#w].Zeit_Abgelaufen THEN
                           IF 4 > #worst_ampel THEN #worst_ampel := 4; END_IF;
                       ELSIF #Bad_Konfig.WT[#w].Vorwarn_Erreicht THEN
                           IF 3 > #worst_ampel THEN #worst_ampel := 3; END_IF;
                       ELSE IF 2 > #worst_ampel THEN #worst_ampel := 2; END_IF;
                       END_IF;
                   ELSE IF 1 > #worst_ampel THEN #worst_ampel := 1; END_IF;
                   END_IF;
               END_IF;
           END_FOR;
       END_IF;
       #Bad_Konfig.Ampel_Status := #worst_ampel;

       //== 10) Ampel-Ausgaenge ==
       #Bad_Konfig.IO_Aus.Ampel_Gruen := FALSE; #Bad_Konfig.IO_Aus.Ampel_Orange := FALSE; #Bad_Konfig.IO_Aus.Ampel_Rot := FALSE;
       CASE #Bad_Konfig.Ampel_Status OF
           0: ; 1: #Bad_Konfig.IO_Aus.Ampel_Gruen := #Blink_Takt;
           2: #Bad_Konfig.IO_Aus.Ampel_Gruen := TRUE;
           3: #Bad_Konfig.IO_Aus.Ampel_Orange := #Blink_Takt;
           4: #Bad_Konfig.IO_Aus.Ampel_Rot := #Blink_Takt;
           5: #Bad_Konfig.IO_Aus.Ampel_Rot := #Blink_Takt;
           6: #Bad_Konfig.IO_Aus.Ampel_Rot := TRUE;
       END_CASE;
       IF #Lampentest THEN
           #Bad_Konfig.IO_Aus.Ampel_Gruen := #Blink_Takt;
           #Bad_Konfig.IO_Aus.Ampel_Orange := #Blink_Takt;
           #Bad_Konfig.IO_Aus.Ampel_Rot := #Blink_Takt;
           #any_hupe := TRUE;
       END_IF;
       #Bad_Konfig.Hupe := #any_hupe;

       //== 11) Peripherie ==
       #Bad_Konfig.IO_Aus.Pumpe := #Bad_Konfig.Ausstattung.HatPumpe AND #Bad_Konfig.Pumpe_Ein AND #hw_ok_ohne_niveau;
       #Bad_Konfig.IO_Aus.Ultraschall_Freigabe := #Bad_Konfig.Ausstattung.HatUltraschall AND #Bad_Konfig.Ultraschall_Ein AND #hw_ok;
       // Pumpe FU: Netzschuetz + Freigabe wenn Sollwert > 0 (ohne Niveau-Pruefung)
       #Bad_Konfig.IO_Aus.Pumpe_FU_Netzschuetz := #Bad_Konfig.Ausstattung.HatPumpe_FU AND (#Bad_Konfig.Pumpe_FU_Soll > 0.0) AND #hw_ok_ohne_niveau;
       #Bad_Konfig.IO_Aus.Pumpe_FU_Freigabe := #Bad_Konfig.IO_Aus.Pumpe_FU_Netzschuetz;

       //== FU-Stoerungen: Fehler nur wenn angesteuert aber nicht bereit (3s Verzoegerung) ==
       #Timer_FU_Pumpe_Stoerung(IN := #Bad_Konfig.IO_Aus.Pumpe_FU_Netzschuetz AND NOT #Bad_Konfig.IO_Ein.FU_Pumpe_Bereit, PT := T#3s);
       #Bad_Konfig.FU_Pumpe_Stoerung := #Timer_FU_Pumpe_Stoerung.Q;

       #Timer_FU_WB1_Stoerung(IN := (#Bad_Konfig.Warenbewegung_Y_Soll > 0.0) AND NOT #Bad_Konfig.IO_Ein.FU_WB1_Bereit, PT := T#3s);
       #Bad_Konfig.FU_WB1_Stoerung := #Timer_FU_WB1_Stoerung.Q;

       #Timer_FU_WB2_Stoerung(IN := (#Bad_Konfig.Warenbewegung_X_Soll > 0.0) AND NOT #Bad_Konfig.IO_Ein.FU_WB2_Bereit, PT := T#3s);
       #Bad_Konfig.FU_WB2_Stoerung := #Timer_FU_WB2_Stoerung.Q;

       //== 12) LEDs ==
       #Bad_Konfig.IO_Aus.LED_Heizung_Aktiv := #irgend_aktiv AND #hw_ok AND NOT #temp_ok;
       #Bad_Konfig.IO_Aus.LED_Stoerung := #irgend_aktiv AND NOT #hw_ok;
       #Bad_Konfig.IO_Aus.LED_Handbetrieb := #hand_aktiv;

       FOR #w := 1 TO 3 DO
           #Bad_Konfig.IO_Aus.LED_Einsetzen[#w] := FALSE;
           IF #Bad_Konfig.WT[#w].Belegt AND NOT #Bad_Konfig.WT[#w].WT_Eingesetzt AND #hw_ok AND #temp_ok THEN
               #Bad_Konfig.IO_Aus.LED_Einsetzen[#w] := #blink[#w];
           END_IF;
       END_FOR;
       FOR #w := 1 TO 3 DO
           #Bad_Konfig.IO_Aus.LED_Entnehmen[#w] := FALSE;
           #Bad_Konfig.IO_Aus.LED_Vorwarn[#w] := FALSE;
           IF #Bad_Konfig.WT[#w].Belegt AND #Bad_Konfig.WT[#w].WT_Eingesetzt THEN
               IF #Bad_Konfig.WT[#w].Zeit_Abgelaufen THEN #Bad_Konfig.IO_Aus.LED_Entnehmen[#w] := #blink[#w];
               ELSIF #Bad_Konfig.WT[#w].Vorwarn_Erreicht THEN
                   #Bad_Konfig.IO_Aus.LED_Entnehmen[#w] := #blink[#w]; #Bad_Konfig.IO_Aus.LED_Vorwarn[#w] := TRUE;
               END_IF;
           END_IF;
       END_FOR;

       //== 13) Prioritaet ==
       #Bad_Konfig.IO_Aus.Prio_Einsetzen_WT := 0;
       FOR #w := 1 TO 3 DO
           IF #Bad_Konfig.WT[#w].Belegt AND NOT #Bad_Konfig.WT[#w].WT_Eingesetzt
              AND #hw_ok AND #temp_ok AND (#Bad_Konfig.IO_Aus.Prio_Einsetzen_WT = 0) THEN
               #Bad_Konfig.IO_Aus.Prio_Einsetzen_WT := #w;
           END_IF;
       END_FOR;
       #Bad_Konfig.IO_Aus.Prio_Entnehmen_WT := 0;
       #ent_prio_rest := T#24h;
       FOR #w := 1 TO 3 DO
           IF #Bad_Konfig.WT[#w].Belegt AND #Bad_Konfig.WT[#w].WT_Eingesetzt AND #Bad_Konfig.WT[#w].Zeit_Abgelaufen THEN
               IF #Bad_Konfig.IO_Aus.Prio_Entnehmen_WT = 0 THEN #Bad_Konfig.IO_Aus.Prio_Entnehmen_WT := #w; END_IF;
           END_IF;
       END_FOR;
       IF #Bad_Konfig.IO_Aus.Prio_Entnehmen_WT = 0 THEN
           FOR #w := 1 TO 3 DO
               IF #Bad_Konfig.WT[#w].Belegt AND #Bad_Konfig.WT[#w].WT_Eingesetzt
                  AND #Bad_Konfig.WT[#w].Vorwarn_Erreicht AND NOT #Bad_Konfig.WT[#w].Zeit_Abgelaufen THEN
                   IF #Bad_Konfig.WT[#w].Restzeit < #ent_prio_rest THEN
                       #ent_prio_rest := #Bad_Konfig.WT[#w].Restzeit;
                       #Bad_Konfig.IO_Aus.Prio_Entnehmen_WT := #w;
                   END_IF;
               END_IF;
           END_FOR;
       END_IF;
END_FUNCTION_BLOCK

FUNCTION_BLOCK "FB_Heizungssteuerung"   // FB11, SCL
{ S7_Optimized_Access := 'TRUE' }
VERSION : 0.1
// stored: AutoNumber true, IsIECCheckEnabled false, IsRetainMemResEnabled false, MemoryReserve 100, SetENOAutomatically false, UDAEnableTagReadback false
   VAR
      Regler_Bad_7 { S7_SetPoint := 'True'} : "FB_Heizungsregelung";
      Regler_Bad_8 { S7_SetPoint := 'True'} : "FB_Heizungsregelung";
      Regler_Bad_12 { S7_SetPoint := 'True'} : "FB_Heizungsregelung";
      Regler_Bad_25_H1 { S7_SetPoint := 'True'} : "FB_Heizungsregelung";
      Regler_Bad_25_H2 { S7_SetPoint := 'True'} : "FB_Heizungsregelung";
      Regler_Bad_36 { S7_SetPoint := 'True'} : "FB_Heizungsregelung";
      Regler_Bad_40 { S7_SetPoint := 'True'} : "FB_Heizungsregelung";
      Regler_Bad_46 { S7_SetPoint := 'True'} : "FB_Heizungsregelung";
   END_VAR
   VAR_TEMP
      sf : Bool;
   END_VAR
BEGIN

       #sf:="DB_Bad_Konfig".Bad_Konfig[7].IO_Ein.FI_Schutz_OK AND "DB_Bad_Konfig".Bad_Konfig[7].IO_Ein.Kein_Uebertemp AND("DB_Bad_Konfig".Bad_Konfig[7].IO_Ein.Niveau_OK OR NOT "DB_Bad_Konfig".Bad_Konfig[7].Ausstattung.HatNiveau);
       #Regler_Bad_7(Soll:="DB_Bad_Konfig".Bad_Konfig[7].Heizung_1_Soll,Ist:="DB_Bad_Konfig".Bad_Konfig[7].Heizung_1_Ist,Freigabe:=#sf);
       "DB_Bad_Konfig".Bad_Konfig[7].IO_Aus.Heizung_1_Regelung:=#Regler_Bad_7.Schuetz;
       "DB_Bad_Konfig".Bad_Konfig[7].IO_Aus.Heizung_1_Sicherheit:=#sf AND("DB_Bad_Konfig".Bad_Konfig[7].Heizung_1_Soll>0.0);
       #sf:="DB_Bad_Konfig".Bad_Konfig[8].IO_Ein.FI_Schutz_OK AND "DB_Bad_Konfig".Bad_Konfig[8].IO_Ein.Kein_Uebertemp AND("DB_Bad_Konfig".Bad_Konfig[8].IO_Ein.Niveau_OK OR NOT "DB_Bad_Konfig".Bad_Konfig[8].Ausstattung.HatNiveau);
       #Regler_Bad_8(Soll:="DB_Bad_Konfig".Bad_Konfig[8].Heizung_1_Soll,Ist:="DB_Bad_Konfig".Bad_Konfig[8].Heizung_1_Ist,Freigabe:=#sf);
       "DB_Bad_Konfig".Bad_Konfig[8].IO_Aus.Heizung_1_Regelung:=#Regler_Bad_8.Schuetz;
       "DB_Bad_Konfig".Bad_Konfig[8].IO_Aus.Heizung_1_Sicherheit:=#sf AND("DB_Bad_Konfig".Bad_Konfig[8].Heizung_1_Soll>0.0);
       #sf:="DB_Bad_Konfig".Bad_Konfig[12].IO_Ein.FI_Schutz_OK AND "DB_Bad_Konfig".Bad_Konfig[12].IO_Ein.Kein_Uebertemp AND("DB_Bad_Konfig".Bad_Konfig[12].IO_Ein.Niveau_OK OR NOT "DB_Bad_Konfig".Bad_Konfig[12].Ausstattung.HatNiveau);
       #Regler_Bad_12(Soll:="DB_Bad_Konfig".Bad_Konfig[12].Heizung_1_Soll,Ist:="DB_Bad_Konfig".Bad_Konfig[12].Heizung_1_Ist,Freigabe:=#sf);
       "DB_Bad_Konfig".Bad_Konfig[12].IO_Aus.Heizung_1_Regelung:=#Regler_Bad_12.Schuetz;
       "DB_Bad_Konfig".Bad_Konfig[12].IO_Aus.Heizung_1_Sicherheit:=#sf AND("DB_Bad_Konfig".Bad_Konfig[12].Heizung_1_Soll>0.0);
       #sf:="DB_Bad_Konfig".Bad_Konfig[25].IO_Ein.FI_Schutz_OK AND "DB_Bad_Konfig".Bad_Konfig[25].IO_Ein.Kein_Uebertemp AND("DB_Bad_Konfig".Bad_Konfig[25].IO_Ein.Niveau_OK OR NOT "DB_Bad_Konfig".Bad_Konfig[25].Ausstattung.HatNiveau);
       #Regler_Bad_25_H1(Soll:="DB_Bad_Konfig".Bad_Konfig[25].Heizung_1_Soll,Ist:="DB_Bad_Konfig".Bad_Konfig[25].Heizung_1_Ist,Freigabe:=#sf);
       "DB_Bad_Konfig".Bad_Konfig[25].IO_Aus.Heizung_1_Regelung:=#Regler_Bad_25_H1.Schuetz;
       #Regler_Bad_25_H2(Soll:="DB_Bad_Konfig".Bad_Konfig[25].Heizung_2_Soll,Ist:="DB_Bad_Konfig".Bad_Konfig[25].Heizung_2_Ist,Freigabe:=#sf);
       "DB_Bad_Konfig".Bad_Konfig[25].IO_Aus.Heizung_2_Regelung:=#Regler_Bad_25_H2.Schuetz;
       "DB_Bad_Konfig".Bad_Konfig[25].IO_Aus.Heizung_1_Sicherheit:=#sf AND(("DB_Bad_Konfig".Bad_Konfig[25].Heizung_1_Soll>0.0)OR("DB_Bad_Konfig".Bad_Konfig[25].Heizung_2_Soll>0.0));
       "DB_Bad_Konfig".Bad_Konfig[25].IO_Aus.Heizung_2_Sicherheit:="DB_Bad_Konfig".Bad_Konfig[25].IO_Aus.Heizung_1_Sicherheit;
       #sf:="DB_Bad_Konfig".Bad_Konfig[36].IO_Ein.FI_Schutz_OK AND "DB_Bad_Konfig".Bad_Konfig[36].IO_Ein.Kein_Uebertemp AND("DB_Bad_Konfig".Bad_Konfig[36].IO_Ein.Niveau_OK OR NOT "DB_Bad_Konfig".Bad_Konfig[36].Ausstattung.HatNiveau);
       #Regler_Bad_36(Soll:="DB_Bad_Konfig".Bad_Konfig[36].Heizung_1_Soll,Ist:="DB_Bad_Konfig".Bad_Konfig[36].Heizung_1_Ist,Freigabe:=#sf);
       "DB_Bad_Konfig".Bad_Konfig[36].IO_Aus.Heizung_1_Regelung:=#Regler_Bad_36.Schuetz;
       "DB_Bad_Konfig".Bad_Konfig[36].IO_Aus.Heizung_1_Sicherheit:=#sf AND("DB_Bad_Konfig".Bad_Konfig[36].Heizung_1_Soll>0.0);
       #sf:="DB_Bad_Konfig".Bad_Konfig[40].IO_Ein.FI_Schutz_OK AND "DB_Bad_Konfig".Bad_Konfig[40].IO_Ein.Kein_Uebertemp AND("DB_Bad_Konfig".Bad_Konfig[40].IO_Ein.Niveau_OK OR NOT "DB_Bad_Konfig".Bad_Konfig[40].Ausstattung.HatNiveau);
       #Regler_Bad_40(Soll:="DB_Bad_Konfig".Bad_Konfig[40].Heizung_1_Soll,Ist:="DB_Bad_Konfig".Bad_Konfig[40].Heizung_1_Ist,Freigabe:=#sf);
       "DB_Bad_Konfig".Bad_Konfig[40].IO_Aus.Heizung_1_Regelung:=#Regler_Bad_40.Schuetz;
       "DB_Bad_Konfig".Bad_Konfig[40].IO_Aus.Heizung_1_Sicherheit:=#sf AND("DB_Bad_Konfig".Bad_Konfig[40].Heizung_1_Soll>0.0);
       #sf:="DB_Bad_Konfig".Bad_Konfig[46].IO_Ein.FI_Schutz_OK AND "DB_Bad_Konfig".Bad_Konfig[46].IO_Ein.Kein_Uebertemp AND("DB_Bad_Konfig".Bad_Konfig[46].IO_Ein.Niveau_OK OR NOT "DB_Bad_Konfig".Bad_Konfig[46].Ausstattung.HatNiveau);
       #Regler_Bad_46(Soll:="DB_Bad_Konfig".Bad_Konfig[46].Heizung_1_Soll,Ist:="DB_Bad_Konfig".Bad_Konfig[46].Heizung_1_Ist,Freigabe:=#sf);
       "DB_Bad_Konfig".Bad_Konfig[46].IO_Aus.Heizung_1_Regelung:=#Regler_Bad_46.Schuetz;
       "DB_Bad_Konfig".Bad_Konfig[46].IO_Aus.Heizung_1_Sicherheit:=#sf AND("DB_Bad_Konfig".Bad_Konfig[46].Heizung_1_Soll>0.0);
END_FUNCTION_BLOCK

FUNCTION_BLOCK "FB_Heizungsregelung"   // FB10, SCL
{ S7_Optimized_Access := 'TRUE' }
VERSION : 0.1
// stored: AutoNumber true, IsIECCheckEnabled false, IsRetainMemResEnabled false, MemoryReserve 100, SetENOAutomatically false, UDAEnableTagReadback false
   VAR_INPUT
      Soll : Real;
      Ist : Real;
      Freigabe : Bool;
   END_VAR
   VAR_OUTPUT
      Schuetz : Bool;
      PT100_Stoerung : Bool;
   END_VAR
   VAR
      Schuetz_Intern : Bool;
   END_VAR
   VAR_TEMP
      einschaltSchwelle : Real;
      ausschaltSchwelle : Real;
   END_VAR
   VAR CONSTANT
      HYSTERESE : Real := 0.2;
      PT100_MIN : Real := -10.0;
      PT100_MAX : Real := 200.0;
   END_VAR
BEGIN

       #PT100_Stoerung:=(#Ist<#PT100_MIN)OR(#Ist>#PT100_MAX);
       IF NOT #Freigabe OR(#Soll<=0.0)OR #PT100_Stoerung THEN #Schuetz_Intern:=FALSE; #Schuetz:=FALSE; RETURN; END_IF;
       #einschaltSchwelle:=#Soll-(#HYSTERESE/2.0); #ausschaltSchwelle:=#Soll+(#HYSTERESE/2.0);
       IF #Ist<#einschaltSchwelle THEN #Schuetz_Intern:=TRUE; ELSIF #Ist>#ausschaltSchwelle THEN #Schuetz_Intern:=FALSE; END_IF;
       #Schuetz:=#Schuetz_Intern;
END_FUNCTION_BLOCK

FUNCTION_BLOCK "FB_FlexKraft"   // FB1, SCL
{ S7_Optimized_Access := 'TRUE' }
VERSION : 0.1
// ==============================================================================
//  FB: Komfort-Wrapper fÃ¼r ein FlexKraft-GerÃ¤t
// ------------------------------------------------------------------------------
//   PflÃ¼ckt das Status-Register in einzelne BOOLs auseinander, baut umgekehrt
//   aus einzelnen BOOLs das Control-Register zusammen und reicht die Sollwerte
//   durch. Es findet KEINE Skalierung statt - der Aufrufer Ã¼bergibt direkt die
//   Modbus-Rohwerte (Spannung in 1/100 V, Strom in 1 A bzw. 0,1 A je HiRes).
// ==============================================================================
// stored: AutoNumber true, IsIECCheckEnabled false, IsRetainMemResEnabled false, MemoryReserve 100, SetENOAutomatically false, UDAEnableTagReadback false
   VAR_INPUT
      bOn : Bool;   // Bit 0 On/Off
      bStartA : Bool;   // Bit 1 Start A
      bBlockA : Bool;   // Bit 2 Block A (Pause)
      bRunProgA : Bool;   // Bit 3 Programm A laufen lassen
      bReverseA : Bool;   // Bit 4 Polung A umkehren
      bReverseB : Bool;   // Bit 5 Polung B umkehren
      bStartB : Bool;   // Bit 7 Start B
      bClrAhA : Bool;   // Bit 8 AhCounter A lÃ¶schen
      bClrAhB : Bool;   // Bit 9 AhCounter B lÃ¶schen
      bClrTimer : Bool;   // Bit 10 ProcessTimer lÃ¶schen
      bBlockB : Bool;   // Bit 12 Block B (Pause)
      bAuxOutA : Bool;   // Bit 13 Auxiliary Out A
      bAuxOutB : Bool;   // Bit 14 Auxiliary Out B
      bRunProgB : Bool;   // Bit 15 Programm B laufen lassen --- Sollwerte (roh, ohne Skalierung) ---
      iSetVoltage_cV : Int;   // Sollspannung 1/100 V (1500 = 15,00 V)
      iSetCurrent_raw : Int;   // Sollstrom 1 A bzw. 0,1 A (siehe HiRes)
      wStartramp_dS : Word;   // Anlauframpe 1/10 s (50 = 5,0 s) --- Bits StatusRegister (Reg 1) ---
   END_VAR
   VAR_OUTPUT
      bAlarm : Bool;   // Bit 0
      bWarning : Bool;   // Bit 1
      bRemote : Bool;   // Bit 2 -> nur wenn TRUE Ã¼bernimmt FK Sollwerte
      bRunningA : Bool;   // Bit 3
      bAhLimitA : Bool;   // Bit 4
      bAhLimitB : Bool;   // Bit 5
      bTimerLimitA : Bool;   // Bit 6
      bVoltageModeA : Bool;   // Bit 7 TRUE = Last zu hochohmig (V-Begrenzung)
      bVoltageModeB : Bool;   // Bit 8
      bUnitOn : Bool;   // Bit 9 (entspricht der grÃ¼nen LED am GerÃ¤t)
      bHiRes : Bool;   // Bit 10 TRUE = Strom in 0,1 A statt 1 A
      bRunningB : Bool;   // Bit 11 --- Istwerte (roh) ---
      iOutVoltage_cV : Int;
      iOutCurrent_raw : Int;   // --- Roh-Bitregister fÃ¼r Detailauswertung in der Applikation ---
      wWarnings : Word;
      wAlarms : Word;
   END_VAR
   VAR_IN_OUT
      stDev : "UDT_FlexKraft_Device";
   END_VAR
BEGIN

   //--------------------------------------------------------------------------
   // 1) Output zusammenbauen
   //--------------------------------------------------------------------------
   #stDev.Out.PageNo := 16#0000;

   #stDev.Out.ControlRegister.%X0 := #bOn;
   #stDev.Out.ControlRegister.%X1 := #bStartA;
   #stDev.Out.ControlRegister.%X2 := #bBlockA;
   #stDev.Out.ControlRegister.%X3 := #bRunProgA;
   #stDev.Out.ControlRegister.%X4 := #bReverseA;
   #stDev.Out.ControlRegister.%X5 := #bReverseB;
   #stDev.Out.ControlRegister.%X6 := FALSE;       // reserviert
   #stDev.Out.ControlRegister.%X7 := #bStartB;
   #stDev.Out.ControlRegister.%X8 := #bClrAhA;
   #stDev.Out.ControlRegister.%X9 := #bClrAhB;
   #stDev.Out.ControlRegister.%X10 := #bClrTimer;
   #stDev.Out.ControlRegister.%X11 := FALSE;       // reserviert
   #stDev.Out.ControlRegister.%X12 := #bBlockB;
   #stDev.Out.ControlRegister.%X13 := #bAuxOutA;
   #stDev.Out.ControlRegister.%X14 := #bAuxOutB;
   #stDev.Out.ControlRegister.%X15 := #bRunProgB;

   #stDev.Out.SetVoltage := #iSetVoltage_cV;
   #stDev.Out.SetCurrent := #iSetCurrent_raw;
   #stDev.Out.Startramp := #wStartramp_dS;

   //--------------------------------------------------------------------------
   // 2) StatusRegister auseinanderpflÃ¼cken
   //--------------------------------------------------------------------------
   #bAlarm := #stDev.In.StatusRegister.%X0;
   #bWarning := #stDev.In.StatusRegister.%X1;
   #bRemote := #stDev.In.StatusRegister.%X2;
   #bRunningA := #stDev.In.StatusRegister.%X3;
   #bAhLimitA := #stDev.In.StatusRegister.%X4;
   #bAhLimitB := #stDev.In.StatusRegister.%X5;
   #bTimerLimitA := #stDev.In.StatusRegister.%X6;
   #bVoltageModeA := #stDev.In.StatusRegister.%X7;
   #bVoltageModeB := #stDev.In.StatusRegister.%X8;
   #bUnitOn := #stDev.In.StatusRegister.%X9;
   #bHiRes := #stDev.In.StatusRegister.%X10;
   #bRunningB := #stDev.In.StatusRegister.%X11;

   //--------------------------------------------------------------------------
   // 3) Istwerte und Roh-Bitregister durchreichen
   //--------------------------------------------------------------------------
   #iOutVoltage_cV := #stDev.In.OutputVoltage;
   #iOutCurrent_raw := #stDev.In.OutputCurrent;
   #wWarnings := #stDev.In.WarningsRegister;
   #wAlarms := #stDev.In.AlarmsRegister;
END_FUNCTION_BLOCK

FUNCTION "FC_Fehlermeldungen" : Void   // FC5, SCL
{ S7_Optimized_Access := 'TRUE' }
VERSION : 0.1
// stored: AutoNumber true, IsIECCheckEnabled false, SetENOAutomatically false, UDAEnableTagReadback false
BEGIN

       // FI-Schutz (invertiert: Eingang TRUE = OK, Fehler = NOT)
       "DB_Fehlermeldungen".FI_Heizung_Bad_7  := NOT "FI-Schutz 200F1 Heizung Bad 7 ist O.K.";
       "DB_Fehlermeldungen".FI_Heizung_Bad_8  := NOT "FI-Schutz 210F1 Heizung Bad 8 ist O.K.";
       "DB_Fehlermeldungen".FI_Heizung_Bad_12 := NOT "FI-Schutz 220F1 Heizung Bad 12 ist O.K.";
       "DB_Fehlermeldungen".FI_Heizung_Bad_25 := NOT ("Motorschutz und FI-Schutz 270Q1, 270F1 Heizung Bad 25 sind O.K." AND "Motorschutz und FI-Schutz 271Q1, 271F1 Heizung Bad 25 sind O.K.");
       "DB_Fehlermeldungen".FI_Heizung_Bad_36 := NOT "FI-Schutz 300F1 Heizung Bad 36 ist O.K.";
       "DB_Fehlermeldungen".FI_Heizung_Bad_40 := NOT "FI-Schutz 310F1 Heizung Bad 40 ist O.K.";
       "DB_Fehlermeldungen".FI_Heizung_Bad_46 := NOT "FI-Schutz 340F1 Heizung Bad 46 ist O.K.";

       // Uebertemperatur (invertiert)
       "DB_Fehlermeldungen".Uebertemp_Bad_7  := NOT "Heizung Bad 7 Keine uebertemperatur";
       "DB_Fehlermeldungen".Uebertemp_Bad_8  := NOT "Heizung Bad 8 Keine uebertemperatur";
       "DB_Fehlermeldungen".Uebertemp_Bad_12 := NOT "Heizung Bad 12 Keine uebertemperatur";
       "DB_Fehlermeldungen".Uebertemp_Bad_25 := NOT "Heizung Bad 25 Keine uebertemperatur";
       "DB_Fehlermeldungen".Uebertemp_Bad_36 := NOT "Heizung Bad 36 Keine uebertemperatur";
       "DB_Fehlermeldungen".Uebertemp_Bad_40 := NOT "Heizung Bad 40 Keine uebertemperatur";
       "DB_Fehlermeldungen".Uebertemp_Bad_46 := NOT "Heizung Bad 46 Keine uebertemperatur";

       // Motorschutz Pumpe (invertiert)
       "DB_Fehlermeldungen".Motorschutz_Pumpe_Bad_8  := NOT "Motorschutz 215Q1 Pumpe Bad 8 ist O.K.";
       "DB_Fehlermeldungen".Motorschutz_Pumpe_Bad_12 := NOT "Motorschutz 225Q1 Pumpe Bad 12 ist O.K.";
       "DB_Fehlermeldungen".Motorschutz_Pumpe_Bad_14 := NOT "Motorschutz 235Q1 Pumpe Bad 14 ist O.K.";
       "DB_Fehlermeldungen".Motorschutz_Pumpe_Bad_18 := NOT "Motorschutz 245Q1 Pumpe Bad 18 ist O.K.";
       "DB_Fehlermeldungen".Motorschutz_Pumpe_Bad_19 := NOT "Motorschutz 255Q1 Pumpe Bad 19 ist O.K.";
       "DB_Fehlermeldungen".Motorschutz_Pumpe_Bad_21 := NOT "Motorschutz 265Q1 Pumpe Bad 21 ist O.K.";
       "DB_Fehlermeldungen".Motorschutz_Pumpe_Bad_25 := NOT "Motorschutz 275Q1 Pumpe Bad 25 ist O.K.";
       "DB_Fehlermeldungen".Motorschutz_Pumpe_Bad_26 := NOT "Motorschutz 285Q1 Pumpe Bad 26 ist O.K.";
       "DB_Fehlermeldungen".Motorschutz_Pumpe_Bad_31 := NOT "Motorschutz 295Q1 Pumpe Bad 31 ist O.K.";
       "DB_Fehlermeldungen".Motorschutz_Pumpe_Bad_41 := NOT "Motorschutz 325Q1 Pumpe Bad 41 ist O.K.";
       "DB_Fehlermeldungen".Motorschutz_Pumpe_Bad_45 := NOT "Motorschutz 335Q1 Pumpe Bad 45 ist O.K.";

       // Wartungsschalter Pumpe (invertiert)
       "DB_Fehlermeldungen".Wartungsschalter_Pumpe_Bad_8  := NOT "Wartungsschalter Pumpe Bad 8 ist eingeschaltet";
       "DB_Fehlermeldungen".Wartungsschalter_Pumpe_Bad_12 := NOT "Wartungsschalter Pumpe Bad 12 ist eingeschaltet";
       "DB_Fehlermeldungen".Wartungsschalter_Pumpe_Bad_14 := NOT "Wartungsschalter Pumpe Bad 14 ist eingeschaltet";
       "DB_Fehlermeldungen".Wartungsschalter_Pumpe_Bad_18 := NOT "Wartungsschalter Pumpe Bad 18 ist eingeschaltet";
       "DB_Fehlermeldungen".Wartungsschalter_Pumpe_Bad_19 := NOT "Wartungsschalter Pumpe Bad 19 ist eingeschaltet";
       "DB_Fehlermeldungen".Wartungsschalter_Pumpe_Bad_21 := NOT "Wartungsschalter Pumpe Bad 21 ist eingeschaltet";
       "DB_Fehlermeldungen".Wartungsschalter_Pumpe_Bad_25 := NOT "Wartungsschalter Pumpe Bad 25 ist eingeschaltet";
       "DB_Fehlermeldungen".Wartungsschalter_Pumpe_Bad_26 := NOT "Wartungsschalter Pumpe Bad 26 ist eingeschaltet";
       "DB_Fehlermeldungen".Wartungsschalter_Pumpe_Bad_31 := NOT "Wartungsschalter Pumpe Bad 31 ist eingeschaltet";
       "DB_Fehlermeldungen".Wartungsschalter_Pumpe_Bad_41 := NOT "Wartungsschalter Pumpe Bad 41 ist eingeschaltet";
       "DB_Fehlermeldungen".Wartungsschalter_Pumpe_Bad_45 := NOT "Wartungsschalter Pumpe Bad 45 ist eingeschaltet";

       // Niveau (invertiert)
       "DB_Fehlermeldungen".Niveau_Bad_7  := NOT "Niveau Bad 7 OK";
       "DB_Fehlermeldungen".Niveau_Bad_8  := NOT "Niveau Bad 8 OK";
       "DB_Fehlermeldungen".Niveau_Bad_12 := NOT "Niveau Bad 12 OK";
       "DB_Fehlermeldungen".Niveau_Bad_25 := NOT "Niveau Bad 25 OK";
       "DB_Fehlermeldungen".Niveau_Bad_36 := NOT "Niveau Bad 36 OK";
       "DB_Fehlermeldungen".Niveau_Bad_40 := NOT "Niveau Bad 40 OK";
       "DB_Fehlermeldungen".Niveau_Bad_46 := NOT "Niveau Bad 46 OK";

       // FU Stoerung (aus FB_Bad, 3s verzoegert: angesteuert aber nicht bereit)
       "DB_Fehlermeldungen".FU_Pumpe_Bad_25 := "DB_Bad_Konfig".Bad_Konfig[25].FU_Pumpe_Stoerung;
       "DB_Fehlermeldungen".FU_WB1_Bad_25   := "DB_Bad_Konfig".Bad_Konfig[25].FU_WB1_Stoerung;
       "DB_Fehlermeldungen".FU_WB2_Bad_25   := "DB_Bad_Konfig".Bad_Konfig[25].FU_WB2_Stoerung;

       // Motorschutz Warenbewegung (invertiert)
       "DB_Fehlermeldungen".Motorschutz_WB1_Bad_25 := NOT "Motorschutz 276Q1 Warenbewegung 1 Bad 25 ist O.K.";
       "DB_Fehlermeldungen".Motorschutz_WB2_Bad_25 := NOT "Motorschutz 277Q1 Warenbewegung 2 Bad 25 ist O.K.";

       // PT100 Sensorstoerung (direkt aus Heizungsregelung)
       "DB_Fehlermeldungen".PT100_Bad_7     := "FB_Anlagensteuerung_DB".Heizung.Regler_Bad_7.PT100_Stoerung;
       "DB_Fehlermeldungen".PT100_Bad_8     := "FB_Anlagensteuerung_DB".Heizung.Regler_Bad_8.PT100_Stoerung;
       "DB_Fehlermeldungen".PT100_Bad_12    := "FB_Anlagensteuerung_DB".Heizung.Regler_Bad_12.PT100_Stoerung;
       "DB_Fehlermeldungen".PT100_Bad_25_H1 := "FB_Anlagensteuerung_DB".Heizung.Regler_Bad_25_H1.PT100_Stoerung;
       "DB_Fehlermeldungen".PT100_Bad_25_H2 := "FB_Anlagensteuerung_DB".Heizung.Regler_Bad_25_H2.PT100_Stoerung;
       "DB_Fehlermeldungen".PT100_Bad_36    := "FB_Anlagensteuerung_DB".Heizung.Regler_Bad_36.PT100_Stoerung;
       "DB_Fehlermeldungen".PT100_Bad_40    := "FB_Anlagensteuerung_DB".Heizung.Regler_Bad_40.PT100_Stoerung;
       "DB_Fehlermeldungen".PT100_Bad_46    := "FB_Anlagensteuerung_DB".Heizung.Regler_Bad_46.PT100_Stoerung;

       // Walchem Controller (TRUE = Alarm, keine Invertierung)
       "DB_Fehlermeldungen".Fehler_Walchem_Controller := "Alarm Walchem Controller";

       // Not-Halt
       "DB_Fehlermeldungen".Not_Halt := NOT "Not-Aus ist OK";
END_FUNCTION

FUNCTION "FC_IO_Mapping" : Void   // FC3, SCL
{ S7_Optimized_Access := 'TRUE' }
VERSION : 0.9
// stored: AutoNumber true, IsIECCheckEnabled false, SetENOAutomatically false, UDAEnableTagReadback false
   VAR_INPUT
      Richtung : Int;
   END_VAR
   VAR_TEMP
      "b" : Int;
      w : Int;
      pw : Int;
      hupe_sammel : Bool;
      rawWord : Word;
      rawInt : Int;
   END_VAR
BEGIN

   IF #Richtung = 1 THEN
       FOR #b := 1 TO "c_Anzahl_Bad" DO
           FOR #w := 1 TO 3 DO
               "DB_Bad_Konfig".Bad_Konfig[#b].IO_Ein.WT_Einsetzen[#w] := FALSE;
               "DB_Bad_Konfig".Bad_Konfig[#b].IO_Ein.WT_Entnehmen[#w] := FALSE;
           END_FOR;
       END_FOR;

       // Bad 2, 20, 47: Virtuelle Tasten vom IPC (kein KP8-Modul)
       FOR #w := 1 TO 3 DO
           "DB_Bad_Konfig".Bad_Konfig[2].IO_Ein.WT_Einsetzen[#w] := "DB_IPC_to_CPU".Virtuelle_Tasten.Bad_2.WT_Einsetzen[#w];
           "DB_Bad_Konfig".Bad_Konfig[2].IO_Ein.WT_Entnehmen[#w] := "DB_IPC_to_CPU".Virtuelle_Tasten.Bad_2.WT_Entnehmen[#w];
           "DB_Bad_Konfig".Bad_Konfig[20].IO_Ein.WT_Einsetzen[#w] := "DB_IPC_to_CPU".Virtuelle_Tasten.Bad_20.WT_Einsetzen[#w];
           "DB_Bad_Konfig".Bad_Konfig[20].IO_Ein.WT_Entnehmen[#w] := "DB_IPC_to_CPU".Virtuelle_Tasten.Bad_20.WT_Entnehmen[#w];
           "DB_Bad_Konfig".Bad_Konfig[47].IO_Ein.WT_Einsetzen[#w] := "DB_IPC_to_CPU".Virtuelle_Tasten.Bad_47.WT_Einsetzen[#w];
           "DB_Bad_Konfig".Bad_Konfig[47].IO_Ein.WT_Entnehmen[#w] := "DB_IPC_to_CPU".Virtuelle_Tasten.Bad_47.WT_Entnehmen[#w];
       END_FOR;

